(* IEC 61131-3 sources: ZPLC/conformance/cmp (part 2) *)

(* ---- cmp-020-two-enums-same-value-name.st ---- *)
TYPE A : (X, Y); END_TYPE
TYPE B : (Y, Z); END_TYPE

PROGRAM Main
VAR
  fromA AT %QW0 : INT;
  fromB AT %QW1 : INT;
  zB AT %QW2 : INT;
END_VAR
  fromA := A#Y;
  fromB := B#Y;
  zB := B#Z;
END_PROGRAM

(* ---- cmp-021-concat-leaves-its-arguments.st ---- *)
PROGRAM Main
VAR
  a : STRING[16] := 'ab';
  b : STRING[16] := 'cd';
  r : STRING[16];
  la AT %QW0 : INT;
  lb AT %QW1 : INT;
  lr AT %QW2 : INT;
  ok AT %QX6.0 : BOOL;
END_VAR
  r := CONCAT(a, b);
  la := LEN(a);
  lb := LEN(b);
  lr := LEN(r);
  ok := r = 'abcd';
END_PROGRAM

(* ---- cmp-021-find.st ---- *)
PROGRAM Main
VAR
  s : STRING[16] := 'HELLO';
  p1 AT %QW0 : INT;
  p2 AT %QW1 : INT;
  p3 AT %QW2 : INT;
  p4 AT %QW3 : INT;
END_VAR
  p1 := FIND(s, 'LL');
  p2 := FIND(s, 'H');
  p3 := FIND(s, 'LOL');
  p4 := FIND(s, 'O');
END_PROGRAM

(* ---- cmp-021-function-returning-a-string.st ---- *)
FUNCTION Tag : STRING[8]
VAR_INPUT n : INT; END_VAR
  IF n = 1 THEN
    Tag := 'one';
  ELSE
    Tag := 'other';
  END_IF;
END_FUNCTION

PROGRAM Main
VAR
  r : STRING[12];
  l AT %QW0 : INT;
  ok AT %QX2.0 : BOOL;
END_VAR
  r := CONCAT(Tag(1), Tag(2));
  l := LEN(r);
  ok := r = 'oneother';
END_PROGRAM

(* ---- cmp-021-initial-literal-longer-than-capacity-rejected.st ---- *)
PROGRAM Main
VAR
  s : STRING[3] := 'abcd';
END_VAR
END_PROGRAM

(* ---- cmp-021-insert-delete-replace.st ---- *)
PROGRAM Main
VAR
  s : STRING[16] := 'HELLO';
  i : STRING[16];
  d : STRING[16];
  r : STRING[16];
  ls AT %QW0 : INT;
  oki AT %QX2.0 : BOOL;
  okd AT %QX2.1 : BOOL;
  okr AT %QX2.2 : BOOL;
END_VAR
  i := INSERT(s, 'XY', 2);
  d := DELETE(s, 2, 2);
  r := REPLACE(s, 'AB', 2, 3);
  ls := LEN(s);
  oki := i = 'HEXYLLO';
  okd := d = 'HLO';
  okr := r = 'HABO';
END_PROGRAM

(* ---- cmp-021-left-and-right-beyond-the-length.st ---- *)
PROGRAM Main
VAR
  s : STRING[16] := 'abc';
  l : STRING[16];
  r : STRING[16];
  ll AT %QW0 : INT;
  lr AT %QW1 : INT;
  z AT %QW2 : INT;
END_VAR
  l := LEFT(s, 10);
  r := RIGHT(s, 10);
  ll := LEN(l);
  lr := LEN(r);
  z := LEN(LEFT(s, 0));
END_PROGRAM

(* ---- cmp-021-left-right-mid-keep-the-argument.st ---- *)
PROGRAM Main
VAR
  s : STRING[16] := 'HELLO';
  l : STRING[16];
  r : STRING[16];
  m : STRING[16];
  ls AT %QW0 : INT;
  okl AT %QX2.0 : BOOL;
  okr AT %QX2.1 : BOOL;
  okm AT %QX2.2 : BOOL;
END_VAR
  l := LEFT(s, 2);
  r := RIGHT(s, 3);
  m := MID(s, 2, 3);
  ls := LEN(s);
  okl := l = 'HE';
  okr := r = 'LLO';
  okm := m = 'ELL';
END_PROGRAM

(* ---- cmp-021-literal-longer-than-capacity-rejected.st ---- *)
PROGRAM Main
VAR
  s : STRING[3];
END_VAR
  s := 'abcd';
END_PROGRAM

(* ---- cmp-021-nested-string-functions.st ---- *)
PROGRAM Main
VAR
  a : STRING[16] := 'one';
  b : STRING[16] := 'two';
  r : STRING[16];
  l AT %QW0 : INT;
  ok AT %QX2.0 : BOOL;
  eq AT %QX2.1 : BOOL;
END_VAR
  r := CONCAT(LEFT(a, 2), RIGHT(b, 2));
  l := LEN(r);
  ok := r = 'onwo';
  eq := LEFT(a, 1) = LEFT('ozone', 1);
END_PROGRAM

(* ---- cmp-021-string-assign-length.st ---- *)
PROGRAM Text
VAR
  s : STRING;
  n AT %QW0 : INT;
END_VAR
  s := 'hello';
  n := LEN(s);
END_PROGRAM

(* ---- cmp-021-string-assignment-between-variables.st ---- *)
PROGRAM Main
VAR
  a : STRING[16];
  b : STRING[16];
  la AT %QW0 : INT;
  lb AT %QW1 : INT;
  same AT %QX4.0 : BOOL;
END_VAR
  a := 'hello';
  b := a;
  a := 'x';
  la := LEN(a);
  lb := LEN(b);
  same := b = 'hello';
END_PROGRAM

(* ---- cmp-021-string-buffer-survives-a-function-call.st ---- *)
FUNCTION Mark : INT
VAR_INPUT k : INT; END_VAR
  Mark := LEN(CONCAT('abc', 'defg')) + k;
END_FUNCTION

FUNCTION Pair : INT
VAR_INPUT
  x : STRING[8];
  m : INT;
END_VAR
  Pair := LEN(x) * 100 + m;
END_FUNCTION

PROGRAM Main
VAR
  a : STRING[8] := 'hello';
  r AT %QW0 : INT;
END_VAR
  r := Pair(LEFT(a, 2), Mark(1));
END_PROGRAM

(* ---- cmp-021-string-built-from-itself.st ---- *)
PROGRAM Main
VAR
  e : STRING[8] := 'AB';
  f : STRING[8] := 'AB';
  g : STRING[8] := 'ABCD';
  h : STRING[8] := 'ABCDE';
  okE AT %QX0.0 : BOOL;
  okF AT %QX0.1 : BOOL;
  okG AT %QX0.2 : BOOL;
  okH AT %QX0.3 : BOOL;
END_VAR
  e := CONCAT(e, e);
  f := CONCAT('xy', f);
  g := INSERT(g, '--', 2);
  h := REPLACE(h, 'Y', 2, 3);
  okE := e = 'ABAB';
  okF := f = 'xyAB';
  okG := g = 'AB--CD';
  okH := h = 'AYE';
END_PROGRAM

(* ---- cmp-021-string-comparison.st ---- *)
PROGRAM Main
VAR
  a : STRING[16] := 'abc';
  b : STRING[16] := 'abc';
  c : STRING[16] := 'abd';
  same AT %QX0.0 : BOOL;
  differ AT %QX0.1 : BOOL;
  literal AT %QX0.2 : BOOL;
END_VAR
  same := a = b;
  differ := a <> c;
  literal := c = 'abd';
END_PROGRAM

(* ---- cmp-021-string-cut-in-place.st ---- *)
PROGRAM Main
VAR
  a : STRING[8] := 'ABCDEFGH';
  b : STRING[8] := 'ABCDEFGH';
  c : STRING[8] := 'ABCDEFGH';
  d : STRING[8] := 'ABCDEFGH';
  okA AT %QX0.0 : BOOL;
  okB AT %QX0.1 : BOOL;
  okC AT %QX0.2 : BOOL;
  okD AT %QX0.3 : BOOL;
  lenA AT %QW1 : INT;
END_VAR
  a := LEFT(a, 3);
  b := RIGHT(b, 3);
  c := MID(c, 3, 2);
  d := DELETE(d, 3, 4);
  okA := a = 'ABC';
  okB := b = 'FGH';
  okC := c = 'CD';
  okD := d = 'ABGH';
  lenA := LEN(a);
END_PROGRAM

(* ---- cmp-021-string-function-into-array-element.st ---- *)
PROGRAM Main
VAR
  names : ARRAY[0..2] OF STRING[10];
  i : INT := 1;
  src : STRING[10] := 'pressure';
  l AT %QW0 : INT;
  ok AT %QX2.0 : BOOL;
END_VAR
  names[i] := LEFT(src, 4);
  l := LEN(names[1]);
  ok := names[1] = 'pres';
END_PROGRAM

(* ---- cmp-021-string-function-keeps-argument.st ---- *)
PROGRAM Text
VAR
  left AT %QW0 : INT;
  whole AT %QW1 : INT;
END_VAR
  left := LEN(LEFT('hello', 2));
  whole := LEN('hello');
END_PROGRAM

(* ---- cmp-021-string-function-reading-its-target-in-a-count.st ---- *)
PROGRAM Main
VAR
  k : STRING[8] := 'abcdef';
  t : STRING[8] := 'wxyz';
  okK AT %QX0.0 : BOOL;
  okT AT %QX0.1 : BOOL;
END_VAR
  k := LEFT(k, LEN(k) - 2);
  t := LEFT(t, LEN(k) - 1);
  okK := k = 'abcd';
  okT := t = 'wxy';
END_PROGRAM

(* ---- cmp-021-string-initial-values.st ---- *)
PROGRAM Main
VAR
  a : STRING := 'abc';
  b : STRING[10] := 'hi';
  c : STRING[16];
  la AT %QW0 : INT;
  lb AT %QW1 : INT;
  lc AT %QW2 : INT;
  ok AT %QX6.0 : BOOL;
END_VAR
  la := LEN(a);
  lb := LEN(b);
  lc := LEN(c);
  ok := b = 'hi';
END_PROGRAM

(* ---- cmp-021-string-literal-length.st ---- *)
PROGRAM Text
VAR
  n AT %QW0 : INT;
END_VAR
  n := LEN('hello');
END_PROGRAM

(* ---- cmp-021-string-members-and-elements.st ---- *)
TYPE Label : STRUCT id : INT; text : STRING[12]; END_STRUCT END_TYPE

PROGRAM Main
VAR
  l : Label;
  a : ARRAY[0..1] OF STRING[8];
  lt AT %QW0 : INT;
  la AT %QW1 : INT;
  id AT %QW2 : INT;
  ok AT %QX6.0 : BOOL;
END_VAR
  l.id := 42;
  l.text := 'motor 1';
  a[1] := 'pump';
  lt := LEN(l.text);
  la := LEN(a[1]);
  id := l.id;
  ok := a[1] = 'pump';
END_PROGRAM

(* ---- cmp-021-string-parameter-is-a-copy.st ---- *)
FUNCTION Shout : INT
VAR_INPUT text : STRING[16]; END_VAR
  text := CONCAT(text, '!');
  Shout := LEN(text);
END_FUNCTION

PROGRAM Main
VAR
  s : STRING[16] := 'hello';
  inside AT %QW0 : INT;
  outside AT %QW1 : INT;
END_VAR
  inside := Shout(s);
  outside := LEN(s);
END_PROGRAM

(* ---- cmp-021-string-truncates-to-its-capacity.st ---- *)
PROGRAM Main
VAR
  long : STRING[16] := 'abcdefgh';
  short : STRING[5];
  l AT %QW0 : INT;
  ok AT %QX2.0 : BOOL;
END_VAR
  short := long;
  l := LEN(short);
  ok := short = 'abcde';
END_PROGRAM

(* ---- cmp-021-string-with-capacity.st ---- *)
PROGRAM Text
VAR
  s : STRING[20];
  n AT %QW0 : INT;
END_VAR
  s := 'hello';
  n := LEN(s);
END_PROGRAM

(* ---- cmp-021-wstring-assignment.st ---- *)
PROGRAM Main
VAR
  a : WSTRING[10] := "hi";
  b : WSTRING[10];
  la AT %QW0 : INT;
  lb AT %QW1 : INT;
END_VAR
  b := "world";
  la := LEN(a);
  lb := LEN(b);
  a := b;
  la := LEN(a) * 10 + la;
END_PROGRAM

(* ---- cmp-021-wstring-literal-length.st ---- *)
PROGRAM WideLiteral
VAR
  n AT %QW0 : INT;
END_VAR
  n := LEN("abcd");
END_PROGRAM

(* ---- cmp-021-wstring-variable-length.st ---- *)
PROGRAM WideVariable
VAR
  w : WSTRING := "abcd";
  n AT %QW0 : INT;
END_VAR
  n := LEN(w);
END_PROGRAM

(* ---- cmp-022-array-bound-constant-expression.st ---- *)
VAR_GLOBAL CONSTANT N : INT := 2; END_VAR

PROGRAM Main
VAR
  a : ARRAY[N - 2 .. N * 2 - 1] OF INT;
  last AT %QW0 : INT;
END_VAR
  a[3] := 33;
  last := a[3];
END_PROGRAM

(* ---- cmp-022-array-constant-bound.st ---- *)
VAR_GLOBAL CONSTANT N : INT := 4; END_VAR

PROGRAM Table
VAR
  a : ARRAY[0..N] OF INT;
  last AT %QW0 : INT;
END_VAR
  a[4] := 9;
  last := a[4];
END_PROGRAM

(* ---- cmp-022-array-element-read-write.st ---- *)
PROGRAM Table
VAR
  a : ARRAY[1..4] OF INT;
  i : INT;
  third AT %QW0 : INT;
END_VAR
  FOR i := 1 TO 4 DO
    a[i] := i * 10;
  END_FOR;
  third := a[3];
END_PROGRAM

(* ---- cmp-022-array-index-from-array.st ---- *)
PROGRAM Main
VAR
  b : ARRAY[0..2] OF INT;
  a : ARRAY[0..4] OF DINT;
  v AT %QD0 : DINT;
END_VAR
  b[1] := 4;
  a[4] := 654321;
  v := a[b[1]];
END_PROGRAM

(* ---- cmp-022-array-initialiser-large-repeat.st ---- *)
PROGRAM Main
VAR
  a : ARRAY[0..99] OF INT := [100(3)];
  first AT %QW0 : INT;
  last AT %QW1 : INT;
  after AT %QW2 : INT;
END_VAR
  first := a[0];
  last := a[99];
  after := a[50] + 4;
END_PROGRAM

(* ---- cmp-022-array-initialiser-list.st ---- *)
PROGRAM Table
VAR
  a : ARRAY[0..2] OF INT := [1, 2, 3];
  seen AT %QW0 : INT;
END_VAR
  seen := a[1];
END_PROGRAM

(* ---- cmp-022-array-initialiser-of-structures.st ---- *)
TYPE Pt : STRUCT x : INT; z : DINT; END_STRUCT END_TYPE

PROGRAM Main
VAR
  a : ARRAY[0..1] OF Pt := [(x := 1, z := 100000), (x := 2, z := 200000)];
  x1 AT %QW0 : INT;
  z0 AT %QD1 : DINT;
  z1 AT %QD2 : DINT;
END_VAR
  x1 := a[1].x;
  z0 := a[0].z;
  z1 := a[1].z;
END_PROGRAM

(* ---- cmp-022-array-initialiser-repeat.st ---- *)
PROGRAM Table
VAR
  a : ARRAY[0..3] OF INT := [4(7)];
  seen AT %QW0 : INT;
END_VAR
  seen := a[3];
END_PROGRAM

(* ---- cmp-022-array-initialiser-two-dimensions.st ---- *)
PROGRAM Main
VAR
  a : ARRAY[0..1, 0..2] OF INT := [[1, 2, 3], [4, 5, 6]];
  b : ARRAY[0..1, 0..1] OF INT := [10, 20, 30, 40];
  mid AT %QW0 : INT;
  last AT %QW1 : INT;
  flat AT %QW2 : INT;
END_VAR
  mid := a[1, 1];
  last := a[1, 2];
  flat := b[1, 0];
END_PROGRAM

(* ---- cmp-022-array-inside-structure.st ---- *)
TYPE Rec : STRUCT n : INT; a : ARRAY[1..3] OF DINT; tail : INT; END_STRUCT END_TYPE

PROGRAM Main
VAR
  s : Rec;
  i : INT;
  second AT %QD0 : DINT;
  tail AT %QW2 : INT;
END_VAR
  s.tail := 77;
  FOR i := 1 TO 3 DO
    s.a[i] := i * 100000;
  END_FOR;
  second := s.a[2];
  tail := s.tail;
END_PROGRAM

(* ---- cmp-022-array-negative-lower-bound.st ---- *)
PROGRAM Table
VAR
  a : ARRAY[-5..5] OF INT;
  total AT %QW0 : INT;
END_VAR
  a[-5] := 3;
  a[0] := 4;
  total := a[-5] + a[0];
END_PROGRAM

(* ---- cmp-022-array-of-lint-negative.st ---- *)
PROGRAM Main
VAR
  a : ARRAY[0..3] OF LINT;
  b : LINT;
  same AT %QX0.0 : BOOL;
  negative AT %QX0.1 : BOOL;
  neighbour AT %QX0.2 : BOOL;
END_VAR
  a[1] := -5;
  a[2] := 7;
  b := a[1];
  same := a[1] = -5;
  negative := b < 0;
  neighbour := a[2] = 7;
END_PROGRAM

(* ---- cmp-022-array-of-lint-variable-index.st ---- *)
PROGRAM Main
VAR
  a : ARRAY[0..3] OF LINT;
  i : INT := 2;
  big : LINT := 5000000000;
  back : LINT;
  same AT %QX0.0 : BOOL;
  other AT %QX0.1 : BOOL;
  low AT %QD1 : DINT;
END_VAR
  a[i] := big;
  a[i + 1] := -9;
  back := a[i];
  same := back = 5000000000;
  other := a[3] = -9;
  low := a[2] - 5000000000;
END_PROGRAM

(* ---- cmp-022-array-of-lint.st ---- *)
PROGRAM Table
VAR
  a : ARRAY[0..3] OF LINT;
  ok AT %QX0.0 : BOOL;
END_VAR
  a[2] := 1;
  ok := a[2] = 1;
END_PROGRAM

(* ---- cmp-022-array-of-real-and-bool.st ---- *)
PROGRAM Main
VAR
  r : ARRAY[0..2] OF REAL;
  f : ARRAY[0..2] OF BOOL;
  sum AT %QD0 : REAL;
  second AT %QX4.0 : BOOL;
  third AT %QX4.1 : BOOL;
END_VAR
  r[0] := 1.5;
  r[1] := 2.25;
  r[2] := 0.25;
  f[1] := TRUE;
  sum := r[0] + r[1] + r[2];
  second := f[1];
  third := f[2];
END_PROGRAM

(* ---- cmp-022-array-of-structures-index-expression.st ---- *)
TYPE Pt : STRUCT x : INT; z : DINT; END_STRUCT END_TYPE

PROGRAM Main
VAR
  a : ARRAY[0..3] OF Pt;
  i : INT;
  z2 AT %QD0 : DINT;
  x3 AT %QW2 : INT;
  x0 AT %QW3 : INT;
END_VAR
  FOR i := 0 TO 3 DO
    a[i].z := i * 1000 + 70000;
    a[i].x := -i;
  END_FOR;
  z2 := a[2].z;
  x3 := a[3].x;
  x0 := a[0].x;
END_PROGRAM

(* ---- cmp-022-array-of-structures.st ---- *)
TYPE Pt : STRUCT x : INT; y : INT; z : DINT; END_STRUCT END_TYPE

PROGRAM Table
VAR
  a : ARRAY[0..3] OF Pt;
  seen AT %QW0 : INT;
END_VAR
  a[1].x := 5;
  seen := a[1].x;
END_PROGRAM

(* ---- cmp-022-array-two-dimensions-negative-bounds.st ---- *)
PROGRAM Main
VAR
  a : ARRAY[-1..1, 0..2] OF INT;
  r : INT;
  c : INT;
  low AT %QW0 : INT;
  high AT %QW1 : INT;
  mid AT %QW2 : INT;
END_VAR
  FOR r := -1 TO 1 DO
    FOR c := 0 TO 2 DO
      a[r, c] := r * 10 + c;
    END_FOR;
  END_FOR;
  low := a[-1, 2];
  high := a[1, 0];
  mid := a[0, 1];
END_PROGRAM

(* ---- cmp-022-multi-dimensional-arrays.st ---- *)
PROGRAM Grid
VAR
  plane : ARRAY[0..1, 0..2] OF INT;
  cube : ARRAY[1..2, 1..2, 1..2] OF DINT;
  gains : ARRAY[0..2] OF REAL;
  flags : ARRAY[0..3] OF BOOL;
  i : INT;
  j : INT;
  corner AT %QW0 : INT;
  inner AT %QW1 : INT;
  far AT %QD1 : DINT;
  gain AT %QD2 : REAL;
  flag AT %QX12.0 : BOOL;
  clear AT %QX12.1 : BOOL;
END_VAR
  FOR i := 0 TO 1 DO
    FOR j := 0 TO 2 DO
      plane[i, j] := i * 10 + j;
    END_FOR;
  END_FOR;
  cube[2, 1, 2] := 212;
  gains[2] := 1.5;
  flags[3] := TRUE;
  corner := plane[1, 2];
  inner := plane[0, 1];
  far := cube[2, 1, 2];
  gain := gains[2];
  flag := flags[3];
  clear := flags[0];
END_PROGRAM

(* ---- cmp-023-array-index-out-of-bounds-faults.st ---- *)
PROGRAM Table
VAR
  a : ARRAY[0..1] OF INT;
  index : INT := 2;
END_VAR
  a[index] := 77;
END_PROGRAM

(* ---- cmp-023-constant-index-in-second-dimension-rejected.st ---- *)
PROGRAM Main
VAR
  a : ARRAY[0..1, 0..2] OF INT;
  v AT %QW0 : INT;
END_VAR
  v := a[1, 3];
END_PROGRAM

(* ---- cmp-023-constant-index-out-of-bounds.st ---- *)
PROGRAM Table
VAR
  a : ARRAY[0..3] OF INT;
END_VAR
  a[10] := 1;
END_PROGRAM

(* ---- cmp-023-index-at-both-bounds-is-accepted.st ---- *)
PROGRAM Main
VAR
  a : ARRAY[2..4] OF INT;
  i : INT;
  first AT %QW0 : INT;
  last AT %QW1 : INT;
END_VAR
  i := 2;
  a[i] := 12;
  i := 4;
  a[i] := 14;
  i := 2;
  first := a[i];
  i := 4;
  last := a[i];
END_PROGRAM

(* ---- cmp-023-index-below-lower-bound-faults.st ---- *)
PROGRAM Main
VAR
  a : ARRAY[2..4] OF INT;
  i : INT := 1;
END_VAR
  a[i] := 5;
END_PROGRAM

(* ---- cmp-023-negative-constant-index-rejected.st ---- *)
PROGRAM Main
VAR
  a : ARRAY[0..3] OF INT;
END_VAR
  a[-1] := 1;
END_PROGRAM

(* ---- cmp-023-read-out-of-bounds-faults.st ---- *)
PROGRAM Main
VAR
  a : ARRAY[0..3] OF DINT;
  i : INT := 4;
  v AT %QD0 : DINT;
END_VAR
  v := a[i];
END_PROGRAM

(* ---- cmp-023-second-dimension-out-of-bounds-faults.st ---- *)
PROGRAM Main
VAR
  a : ARRAY[0..1, 0..2] OF INT;
  j : INT := 3;
  v AT %QW0 : INT;
END_VAR
  v := a[1, j];
END_PROGRAM

(* ---- cmp-024-dereference-of-non-reference-rejected.st ---- *)
PROGRAM Main
VAR
  x : INT;
  y : INT;
END_VAR
  y := x^;
END_PROGRAM

(* ---- cmp-024-null-reference-faults.st ---- *)
PROGRAM Pointer
VAR
  p : REF_TO INT;
  seen AT %QW0 : INT;
END_VAR
  seen := p^;
END_PROGRAM

(* ---- cmp-024-ref-of-another-type.st ---- *)
PROGRAM Pointer
VAR
  r : REAL;
  p : REF_TO INT;
END_VAR
  p := REF(r);
END_PROGRAM

(* ---- cmp-024-ref-to-reads-and-writes-the-referenced-variable.st ---- *)
PROGRAM Reference
VAR
  target : INT := 5;
  link : REF_TO INT;
  seen AT %QW0 : INT;
  moved AT %QW1 : INT;
END_VAR
  link := REF(target);
  seen := link^;
  link^ := 42;
  moved := target;
END_PROGRAM

(* ---- cmp-024-reference-is-null-until-assigned.st ---- *)
PROGRAM Main
VAR
  x : INT;
  p : REF_TO INT;
  before AT %QX0.0 : BOOL;
  after AT %QX0.1 : BOOL;
END_VAR
  before := p = NULL;
  p := REF(x);
  after := p = NULL;
END_PROGRAM

(* ---- cmp-024-reference-of-wrong-type-passed-rejected.st ---- *)
FUNCTION Peek : INT
VAR_INPUT r : REF_TO INT; END_VAR
  Peek := r^;
END_FUNCTION

PROGRAM Main
VAR
  d : DINT;
  seen AT %QW0 : INT;
END_VAR
  seen := Peek(REF(d));
END_PROGRAM

(* ---- cmp-024-reference-of-wrong-type-variable-rejected.st ---- *)
PROGRAM Main
VAR
  d : DINT;
  p : REF_TO INT;
END_VAR
  p := REF(d);
END_PROGRAM

(* ---- cmp-024-reference-passed-to-a-function.st ---- *)
FUNCTION Peek : INT
VAR_INPUT r : REF_TO INT; END_VAR
  Peek := r^;
END_FUNCTION

PROGRAM Main
VAR
  v : INT := 41;
  seen AT %QW0 : INT;
END_VAR
  seen := Peek(REF(v)) + 1;
END_PROGRAM

(* ---- cmp-024-reference-read-and-write.st ---- *)
PROGRAM Main
VAR
  x : INT;
  p : REF_TO INT;
  seen AT %QW0 : INT;
  direct AT %QW1 : INT;
END_VAR
  p := REF(x);
  p^ := 7;
  seen := p^;
  direct := x;
END_PROGRAM

(* ---- cmp-024-reference-stored-in-a-number-rejected.st ---- *)
PROGRAM Main
VAR
  d : DINT;
  e : DINT;
END_VAR
  d := REF(e);
END_PROGRAM

(* ---- cmp-024-reference-to-a-structure.st ---- *)
TYPE Pt : STRUCT x : INT; z : DINT; END_STRUCT END_TYPE

PROGRAM Main
VAR
  s : Pt;
  pp : REF_TO Pt;
  x AT %QW0 : INT;
  z AT %QD1 : DINT;
END_VAR
  pp := REF(s);
  pp^.z := 123456;
  pp^.x := -7;
  x := s.x;
  z := pp^.z;
END_PROGRAM

(* ---- cmp-024-reference-to-member-and-element.st ---- *)
TYPE Pt : STRUCT x : INT; z : DINT; END_STRUCT END_TYPE

PROGRAM Main
VAR
  s : Pt;
  a : ARRAY[0..3] OF DINT;
  pz : REF_TO DINT;
  pe : REF_TO DINT;
  z AT %QD0 : DINT;
  e2 AT %QD1 : DINT;
END_VAR
  pz := REF(s.z);
  pz^ := 123456;
  pe := REF(a[2]);
  pe^ := 654321;
  z := s.z;
  e2 := a[2];
END_PROGRAM

(* ---- cmp-025-fifo-default-size-is-eight.st ---- *)
PROGRAM DefaultQueue
VAR
  push AT %IX0.0 : BOOL;
  item AT %ID1 : DINT;
  line : FIFO;
  count AT %QD0 : DINT;
  full AT %QX4.0 : BOOL;
END_VAR
  line(PUSH := push, DATA_IN := item);
  count := line.COUNT;
  full := line.FULL;
END_PROGRAM

(* ---- cmp-025-function-local-initial-value.st ---- *)
FUNCTION Offset : INT
VAR_INPUT a : INT; END_VAR
VAR k : INT := 100; END_VAR
  Offset := a + k;
END_FUNCTION

PROGRAM Locals
VAR
  seen AT %QW0 : INT;
END_VAR
  seen := Offset(1);
END_PROGRAM

(* ---- cmp-025-global-initial-value.st ---- *)
VAR_GLOBAL G : INT := 42; END_VAR

PROGRAM Globals
VAR
  seen AT %QW0 : INT;
END_VAR
  seen := G;
END_PROGRAM

(* ---- cmp-025-global-structure-and-array-initial-values.st ---- *)
TYPE Pt : STRUCT x : INT := 3; z : DINT := 90000; END_STRUCT END_TYPE

VAR_GLOBAL
  g : Pt;
  t : ARRAY[0..2] OF INT := [4, 5, 6];
END_VAR

PROGRAM Main
VAR
  x AT %QW0 : INT;
  z AT %QD1 : DINT;
  t2 AT %QW4 : INT;
END_VAR
  x := g.x;
  z := g.z;
  t2 := t[2];
END_PROGRAM

(* ---- cmp-025-initial-value-is-written-once.st ---- *)
PROGRAM Main
VAR
  n : INT := 5;
  seen AT %QW0 : INT;
END_VAR
  n := n + 1;
  seen := n;
END_PROGRAM

(* ---- cmp-025-initial-values-of-each-type.st ---- *)
PROGRAM Main
VAR
  flag : BOOL := TRUE;
  ratio : REAL := 1.5;
  big : DINT := -70000;
  wait : TIME := T#2s;
  oflag AT %QX0.0 : BOOL;
  oratio AT %QD1 : REAL;
  obig AT %QD2 : DINT;
  owait AT %QD3 : TIME;
END_VAR
  oflag := flag;
  oratio := ratio;
  obig := big;
  owait := wait;
END_PROGRAM

(* ---- cmp-025-lifo-default-size-is-eight.st ---- *)
PROGRAM DefaultStack
VAR
  push AT %IX0.0 : BOOL;
  item AT %ID1 : DINT;
  pile : LIFO;
  count AT %QD0 : DINT;
  full AT %QX4.0 : BOOL;
END_VAR
  pile(PUSH := push, DATA_IN := item);
  count := pile.COUNT;
  full := pile.FULL;
END_PROGRAM

(* ---- cmp-026-assignment-to-a-constant.st ---- *)
VAR_GLOBAL CONSTANT K : INT := 42; END_VAR

PROGRAM Constants
VAR
  x : INT;
END_VAR
  K := 3;
  x := K;
END_PROGRAM

(* ---- cmp-026-constants-of-real-and-integer.st ---- *)
VAR_GLOBAL CONSTANT
  HALF : REAL := 0.5;
  STEP : INT := 4;
END_VAR

PROGRAM Main
VAR
  r AT %QD0 : REAL;
  n AT %QW2 : INT;
END_VAR
  r := HALF * 3.0;
  n := STEP * 3;
END_PROGRAM

(* ---- cmp-026-global-constant-value.st ---- *)
VAR_GLOBAL CONSTANT K : INT := 42; END_VAR

PROGRAM Constants
VAR
  seen AT %QW0 : INT;
END_VAR
  seen := K;
END_PROGRAM

(* ---- cmp-026-var-constant-assignment-rejected.st ---- *)
PROGRAM Main
VAR CONSTANT
  K : INT := 5;
END_VAR
VAR
  x : INT;
END_VAR
  K := 6;
  x := K;
END_PROGRAM

(* ---- cmp-026-var-constant.st ---- *)
PROGRAM Constants
VAR CONSTANT
  K : INT := 5;
END_VAR
VAR
  seen AT %QW0 : INT;
END_VAR
  seen := K;
END_PROGRAM

(* ---- cmp-027-function-local-initial-value-on-every-call.st ---- *)
FUNCTION Step : INT
VAR_INPUT x : INT; END_VAR
VAR k : INT := 10; END_VAR
  k := k + x;
  Step := k;
END_FUNCTION

PROGRAM Main
VAR
  first AT %QW0 : INT;
  second AT %QW1 : INT;
END_VAR
  first := Step(1);
  second := Step(2);
END_PROGRAM

(* ---- cmp-027-function-local-not-retained.st ---- *)
FUNCTION Count : INT
VAR_INPUT x : INT; END_VAR
VAR k : INT; END_VAR
  k := k + 1;
  Count := k;
END_FUNCTION

PROGRAM Calls
VAR
  first AT %QW0 : INT;
  second AT %QW1 : INT;
END_VAR
  first := Count(0);
  second := Count(0);
END_PROGRAM

(* ---- cmp-027-function-local-string-and-array.st ---- *)
FUNCTION Grow : INT
VAR_INPUT n : INT; END_VAR
VAR
  s : STRING[16];
  a : ARRAY[0..2] OF INT;
END_VAR
  a[1] := a[1] + n;
  s := CONCAT(s, 'ab');
  Grow := LEN(s) * 10 + a[1];
END_FUNCTION

PROGRAM Main
VAR
  r AT %QW0 : INT;
END_VAR
  r := Grow(3);
END_PROGRAM

(* ---- cmp-029-non-retain-accepted.st ---- *)
PROGRAM Volatile
VAR NON_RETAIN
  count : INT;
END_VAR
VAR
  seen AT %QW0 : INT;
END_VAR
  count := count + 1;
  seen := count;
END_PROGRAM

(* ---- cmp-029-retain-and-ordinary-variables-together.st ---- *)
PROGRAM Mixed
VAR RETAIN
  kept : DINT;
  flag : BOOL;
END_VAR
VAR
  plain : INT;
  seen AT %QD0 : DINT;
  mark AT %QX4.0 : BOOL;
END_VAR
  kept := kept + 10;
  flag := kept > 15;
  plain := plain + 1;
  seen := kept + plain;
  mark := flag;
END_PROGRAM

(* ---- cmp-029-retain-global-with-initial-value.st ---- *)
VAR_GLOBAL RETAIN
  total : INT := 10;
END_VAR

PROGRAM Totals
VAR
  seen AT %QW0 : INT;
END_VAR
  total := total + 1;
  seen := total;
END_PROGRAM

(* ---- cmp-029-retain-structure-and-string.st ---- *)
TYPE Pair : STRUCT a : INT := 3; b : INT := 4; END_STRUCT END_TYPE

PROGRAM Mixed
VAR RETAIN
  p : Pair;
  s : STRING[10] := 'abc';
  n : INT := 2;
END_VAR
VAR
  sum AT %QW0 : INT;
  len AT %QW2 : INT;
END_VAR
  n := n + 1;
  sum := p.a + p.b + n;
  len := LEN(s);
END_PROGRAM

(* ---- cmp-029-var-global-retain.st ---- *)
VAR_GLOBAL RETAIN
  total : INT;
END_VAR

PROGRAM Totals
VAR
  seen AT %QW0 : INT;
END_VAR
  total := total + 2;
  seen := total;
END_PROGRAM

(* ---- cmp-029-var-non-retain-is-accepted.st ---- *)
PROGRAM Volatile
VAR NON_RETAIN
  x : INT := 5;
END_VAR
VAR
  q AT %QW0 : INT;
END_VAR
  q := x;
END_PROGRAM

(* ---- cmp-029-var-retain-accepted.st ---- *)
PROGRAM Retained
VAR RETAIN
  count : INT;
END_VAR
VAR
  seen AT %QW0 : INT;
END_VAR
  count := count + 1;
  seen := count;
END_PROGRAM

(* ---- cmp-030-alias-default-value.st ---- *)
TYPE Limit : INT := 100; END_TYPE

PROGRAM Defaults
VAR
  a : Limit;
  b : Limit := 7;
  sum AT %QW0 : INT;
END_VAR
  sum := a + b;
END_PROGRAM

(* ---- cmp-030-alias-of-array-and-structure.st ---- *)
TYPE
  Point : STRUCT x : INT; y : INT; END_STRUCT;
  Marker : Point;
  Samples : ARRAY[0..2] OF INT;
END_TYPE

PROGRAM Aliases
VAR
  m : Marker;
  s : Samples;
  total AT %QW0 : INT;
END_VAR
  m.x := 2;
  m.y := 3;
  s[0] := 10;
  s[2] := 20;
  total := m.x + m.y + s[0] + s[2];
END_PROGRAM

(* ---- cmp-030-alias-refers-to-itself.st ---- *)
TYPE A : B; B : A; END_TYPE

PROGRAM Cycle
VAR
  x : A;
END_VAR
END_PROGRAM

(* ---- cmp-030-function-var-output.st ---- *)
FUNCTION Twice : INT
VAR_INPUT a : INT; END_VAR
VAR_OUTPUT o : INT; END_VAR
  o := a;
  Twice := a + a;
END_FUNCTION

PROGRAM Outputs
VAR
  seen AT %QW0 : INT;
END_VAR
  seen := Twice(3);
END_PROGRAM

(* ---- cmp-030-several-names-one-declaration.st ---- *)
PROGRAM Names
VAR
  a, b : INT;
  total AT %QW0 : INT;
END_VAR
  a := 3;
  b := 4;
  total := a + b;
END_PROGRAM

(* ---- cmp-030-several-names-with-initial-value.st ---- *)
PROGRAM Names
VAR
  a, b, c : INT := 4;
  total AT %QW0 : INT;
END_VAR
  total := a + b + c;
END_PROGRAM

(* ---- cmp-030-several-types-one-block.st ---- *)
TYPE
  A : STRUCT v : INT; END_STRUCT;
  B : (R, G);
END_TYPE

PROGRAM Types
VAR
  a : A;
  seen AT %QW0 : INT;
END_VAR
  a.v := 6;
  seen := a.v;
END_PROGRAM

(* ---- cmp-030-type-alias.st ---- *)
TYPE MyInt : INT; END_TYPE

PROGRAM Alias
VAR
  x : MyInt;
  seen AT %QW0 : INT;
END_VAR
  x := 9;
  seen := x;
END_PROGRAM

(* ---- cmp-030-var-external-type-differs.st ---- *)
VAR_GLOBAL G : INT; END_VAR

PROGRAM External
VAR_EXTERNAL G : REAL; END_VAR
VAR
  seen AT %QW0 : INT;
END_VAR
  seen := 1;
END_PROGRAM

(* ---- cmp-030-var-external-without-global.st ---- *)
PROGRAM External
VAR_EXTERNAL Missing : INT; END_VAR
VAR
  seen AT %QW0 : INT;
END_VAR
  seen := Missing;
END_PROGRAM

(* ---- cmp-030-var-external.st ---- *)
VAR_GLOBAL G : INT; END_VAR

PROGRAM External
VAR_EXTERNAL G : INT; END_VAR
VAR
  seen AT %QW0 : INT;
END_VAR
  G := 5;
  seen := G;
END_PROGRAM

(* ---- cmp-030-var-temp-in-program.st ---- *)
PROGRAM Temporary
VAR_TEMP
  k : INT;
END_VAR
VAR
  seen AT %QW0 : INT;
END_VAR
  k := 6;
  seen := k;
END_PROGRAM

(* ---- cmp-031-0x-form-still-works.st ---- *)
PROGRAM Literal
VAR
  seen AT %QW0 : INT;
END_VAR
  seen := 0xFF;
END_PROGRAM

(* ---- cmp-031-base-not-supported.st ---- *)
PROGRAM Literal
VAR
  seen AT %QW0 : INT;
END_VAR
  seen := 3#12;
END_PROGRAM

(* ---- cmp-031-binary-literal.st ---- *)
PROGRAM Literal
VAR
  seen AT %QW0 : INT;
END_VAR
  seen := 2#1010;
END_PROGRAM

(* ---- cmp-031-c-style-hexadecimal-keeps-working.st ---- *)
PROGRAM CStyle
VAR
  n AT %QW0 : INT;
END_VAR
  n := 0xFF;
END_PROGRAM

(* ---- cmp-031-digit-separator.st ---- *)
PROGRAM Literal
VAR
  seen AT %QW0 : INT;
END_VAR
  seen := 1_000;
END_PROGRAM

(* ---- cmp-031-hexadecimal-literal.st ---- *)
PROGRAM Literal
VAR
  seen AT %QW0 : INT;
END_VAR
  seen := 16#FF;
END_PROGRAM

(* ---- cmp-031-negative-based-literal.st ---- *)
PROGRAM Literal
VAR
  seen AT %QW0 : INT;
END_VAR
  seen := -16#10;
END_PROGRAM

(* ---- cmp-031-octal-literal.st ---- *)
PROGRAM Octal
VAR
  n AT %QW0 : INT;
END_VAR
  n := 8#17;
END_PROGRAM

(* ---- cmp-031-separator-in-based-literal.st ---- *)
PROGRAM Literal
VAR
  seen AT %QW0 : INT;
END_VAR
  seen := 2#1111_0000;
END_PROGRAM

(* ---- cmp-031-typed-literal-out-of-range.st ---- *)
PROGRAM Literal
VAR
  seen AT %QW0 : INT;
END_VAR
  seen := SINT#200;
END_PROGRAM

(* ---- cmp-031-typed-literal.st ---- *)
PROGRAM Literal
VAR
  seen AT %QW0 : INT;
END_VAR
  seen := INT#5;
END_PROGRAM

(* ---- cmp-031-typed-literals-of-each-kind.st ---- *)
PROGRAM Literal
VAR
  small AT %QW0 : INT;
  bits AT %QD2 : DWORD;
  flag AT %QX6.0 : BOOL;
  half AT %QD8 : REAL;
END_VAR
  small := SINT#-3 + INT#4;
  bits := DWORD#16#DEAD_BEEF;
  flag := BOOL#TRUE;
  half := REAL#1.5;
END_PROGRAM

(* ---- cmp-032-ampersand-binds-tighter-than-or.st ---- *)
PROGRAM Logic
VAR
  a : BOOL := TRUE;
  b : BOOL := FALSE;
  c : BOOL := FALSE;
  seen AT %QX0.0 : BOOL;
END_VAR
  seen := a OR b & c;
END_PROGRAM

(* ---- cmp-032-ampersand-operator.st ---- *)
PROGRAM Both
VAR
  a : BOOL := TRUE;
  b : BOOL := TRUE;
  both AT %QX0.0 : BOOL;
END_VAR
  both := a & b;
END_PROGRAM

(* ---- cmp-032-bit-access-of-bool-rejected.st ---- *)
PROGRAM Bits
VAR
  f : BOOL;
  seen AT %QX0.0 : BOOL;
END_VAR
  seen := f.0;
END_PROGRAM

(* ---- cmp-032-bit-access.st ---- *)
PROGRAM Bits
VAR
  w : WORD := 1;
  low AT %QX0.0 : BOOL;
END_VAR
  low := w.0;
END_PROGRAM

(* ---- cmp-032-bit-number-out-of-range.st ---- *)
PROGRAM Bits
VAR
  b : BYTE;
  seen AT %QX0.0 : BOOL;
END_VAR
  seen := b.8;
END_PROGRAM

(* ---- cmp-032-bit-of-lword.st ---- *)
PROGRAM Bits
VAR
  l : LWORD;
  low AT %QX0.0 : BOOL;
  high AT %QX0.1 : BOOL;
  other AT %QX0.2 : BOOL;
END_VAR
  l.40 := TRUE;
  low := l.0;
  high := l.40;
  other := l.39;
END_PROGRAM

(* ---- cmp-032-bit-of-member-and-element.st ---- *)
TYPE Status : STRUCT flags : WORD; END_STRUCT END_TYPE

PROGRAM Bits
VAR
  s : Status;
  a : ARRAY[0..1] OF WORD;
  one AT %QX0.0 : BOOL;
  two AT %QX0.1 : BOOL;
END_VAR
  s.flags := 16#0004;
  a[1] := 16#0100;
  one := s.flags.2;
  a[1].0 := TRUE;
  two := a[1].8 AND a[1].0;
END_PROGRAM

(* ---- cmp-032-bit-set-and-clear.st ---- *)
PROGRAM Bits
VAR
  w AT %QW0 : WORD;
END_VAR
  w := 0;
  w.3 := TRUE;
  w.0 := TRUE;
  w.3 := FALSE;
  w.15 := TRUE;
END_PROGRAM

(* ---- cmp-032-bit-write-in-each-width.st ---- *)
PROGRAM Bits
VAR
  b AT %QB0 : BYTE;
  i AT %QW2 : INT;
  d AT %QD4 : DWORD;
END_VAR
  b.7 := TRUE;
  i.15 := TRUE;
  d.31 := TRUE;
  d.0 := TRUE;
END_PROGRAM

(* ---- cmp-032-block-comment.st ---- *)
PROGRAM Comment
VAR
  seen AT %QW0 : INT;
END_VAR
  /* a comment */ seen := 1;
END_PROGRAM

(* ---- cmp-032-comment-delimiters-inside-comments.st ---- *)
PROGRAM Comments
VAR
  seen AT %QW0 : INT;
END_VAR
  (* a /* inside *) seen := 1;
  /* a (* inside */ seen := seen + 1;
  // (* not an opener
  seen := seen + 1; /* trailing */ (* and another *)
END_PROGRAM

(* ---- cmp-032-empty-statement.st ---- *)
PROGRAM Empty
VAR
  seen AT %QW0 : INT;
END_VAR
  seen := 1;;
END_PROGRAM

(* ---- cmp-032-empty-statements-inside-blocks.st ---- *)
PROGRAM Empty
VAR
  seen AT %QW0 : INT;
END_VAR
  ;
  IF TRUE THEN ; seen := 2;; END_IF;;
  CASE seen OF 2: ; seen := seen + 1; END_CASE;
END_PROGRAM

(* ---- cmp-032-exponent-operator.st ---- *)
PROGRAM Power
VAR
  cube AT %QD0 : REAL;
END_VAR
  cube := 2.0 ** 3.0;
END_PROGRAM

(* ---- cmp-032-power-fractional-exponent.st ---- *)
PROGRAM Power
VAR
  d1 : REAL;
  d2 : REAL;
  d3 : REAL;
  d4 : REAL;
  root AT %QX0.0 : BOOL;
  cube AT %QX0.1 : BOOL;
  big AT %QX0.2 : BOOL;
  small AT %QX0.3 : BOOL;
END_VAR
  d1 := 9.0 ** 0.5 - 3.0;
  d2 := 27.0 ** (1.0 / 3.0) - 3.0;
  d3 := 10.0 ** 2.5 / 316.227766 - 1.0;
  d4 := 0.5 ** 1.5 / 0.35355339 - 1.0;
  root := (d1 < 0.0001) AND (d1 > -0.0001);
  cube := (d2 < 0.0001) AND (d2 > -0.0001);
  big := (d3 < 0.00005) AND (d3 > -0.00005);
  small := (d4 < 0.00005) AND (d4 > -0.00005);
END_PROGRAM

(* ---- cmp-032-power-negative-and-zero-exponent.st ---- *)
PROGRAM Power
VAR
  r AT %QD0 : REAL;
  s AT %QD4 : REAL;
  t AT %QD8 : REAL;
END_VAR
  r := 2.0 ** -2.0;
  s := 5.0 ** 0.0;
  t := 0.0 ** 0.0;
END_PROGRAM

(* ---- cmp-032-power-negative-base.st ---- *)
PROGRAM Power
VAR
  r AT %QD0 : REAL;
  s AT %QD4 : REAL;
END_VAR
  r := (-3.0) ** 3.0;
  s := (-2.0) ** 2.0;
END_PROGRAM

(* ---- cmp-032-power-of-integers.st ---- *)
PROGRAM Power
VAR
  a : INT := 2;
  r AT %QD0 : REAL;
  s AT %QD4 : REAL;
END_VAR
  r := 2 ** 10;
  s := a ** 3;
END_PROGRAM

(* ---- cmp-032-power-precedence.st ---- *)
PROGRAM Power
VAR
  r AT %QD0 : REAL;
  s AT %QD4 : REAL;
END_VAR
  r := -2.0 ** 2.0;
  s := 2.0 * 3.0 ** 2.0;
END_PROGRAM

(* ---- cmp-032-power-zero-base-negative-exponent-faults.st ---- *)
PROGRAM Power
VAR
  zero : REAL := 0.0;
  r AT %QD0 : REAL;
END_VAR
  r := zero ** -1.0;
END_PROGRAM

(* ---- cmp-033-library-block-in-lower-case.st ---- *)
PROGRAM Timer
VAR
  t : ton;
  done AT %QX0.0 : BOOL;
END_VAR
  t(IN := TRUE, PT := T#20ms);
  done := t.Q;
END_PROGRAM

(* ---- cmp-033-library-block-name-as-variable.st ---- *)
PROGRAM Names
VAR
  Pulse : BOOL;
  seen AT %QX0.0 : BOOL;
END_VAR
  Pulse := TRUE;
  seen := Pulse;
END_PROGRAM

(* ---- cmp-034-function-does-not-see-a-program-variable.st ---- *)
FUNCTION Peek : INT
VAR_INPUT n : INT; END_VAR
  Peek := n + hidden;
END_FUNCTION

PROGRAM Scopes
VAR
  hidden : INT := 5;
  out AT %QW0 : INT;
END_VAR
  out := Peek(1);
END_PROGRAM

(* ---- cmp-034-function-locals-do-not-clash.st ---- *)
FUNCTION Pick : INT
VAR_INPUT a : INT; b : INT; END_VAR
VAR tmp : INT; END_VAR
  tmp := a;
  Pick := tmp + b;
END_FUNCTION

FUNCTION Mix : INT
VAR_INPUT b : INT; a : INT; END_VAR
VAR tmp : INT; END_VAR
  tmp := a * 10;
  Mix := tmp + b;
END_FUNCTION

PROGRAM Scopes
VAR
  a : INT := 1000;
  tmp : INT := 2000;
  first AT %QW0 : INT;
  second AT %QW1 : INT;
  kept AT %QW2 : INT;
END_VAR
  first := Pick(1, 2);
  second := Mix(1, 2);
  kept := a + tmp;
END_PROGRAM

(* ---- cmp-034-function-reads-a-global.st ---- *)
VAR_GLOBAL
  base : INT := 100;
END_VAR

FUNCTION Offset : INT
VAR_INPUT n : INT; END_VAR
VAR_EXTERNAL base : INT; END_VAR
  Offset := n + base;
END_FUNCTION

PROGRAM Scopes
VAR
  out AT %QW0 : INT;
  other AT %QW1 : INT;
END_VAR
  out := Offset(5);
  other := Offset(n := 6);
END_PROGRAM

(* ---- cmp-034-function-with-loops-and-locals-of-the-same-name.st ---- *)
FUNCTION SumTo : DINT
VAR_INPUT n : INT; END_VAR
VAR i : INT; total : DINT; END_VAR
  FOR i := 1 TO n DO
    total := total + i;
  END_FOR;
  SumTo := total;
END_FUNCTION

FUNCTION SumSquares : DINT
VAR_INPUT n : INT; END_VAR
VAR i : INT; total : DINT; END_VAR
  FOR i := 1 TO n DO
    total := total + i * i;
  END_FOR;
  SumSquares := total;
END_FUNCTION

PROGRAM Loops
VAR
  i : INT := 100;
  total : DINT := 1000;
  sum AT %QD0 : DINT;
  squares AT %QD1 : DINT;
  again AT %QD2 : DINT;
  program_i AT %QW6 : INT;
END_VAR
  sum := SumTo(4);
  squares := SumSquares(3);
  again := SumTo(4);
  program_i := i;
END_PROGRAM

(* ---- cmp-034-parameter-shadows-program-variable.st ---- *)
FUNCTION Succ : INT
VAR_INPUT a : INT; END_VAR
  Succ := a + 1;
END_FUNCTION

PROGRAM Scopes
VAR
  a : INT := 9;
  total AT %QW0 : INT;
END_VAR
  total := Succ(1) + a;
END_PROGRAM

(* ---- cmp-034-same-parameter-name-two-functions.st ---- *)
FUNCTION Succ : INT
VAR_INPUT a : INT; END_VAR
  Succ := a + 1;
END_FUNCTION

FUNCTION Twice : INT
VAR_INPUT a : INT; END_VAR
  Twice := a * 2;
END_FUNCTION

PROGRAM Scopes
VAR
  total AT %QW0 : INT;
END_VAR
  total := Succ(1) + Twice(2);
END_PROGRAM

(* ---- cmp-035-call-statement-runs-the-function.st ---- *)
VAR_GLOBAL
  counter : INT;
END_VAR

FUNCTION Bump : INT
VAR_INPUT amount : INT; END_VAR
VAR_EXTERNAL counter : INT; END_VAR
  counter := counter + amount;
  Bump := counter;
END_FUNCTION

PROGRAM Statement
VAR
  seen AT %QW0 : INT;
END_VAR
  Bump(2);
  Bump(amount := 3);
  seen := counter;
END_PROGRAM

(* ---- cmp-035-function-call-as-statement.st ---- *)
FUNCTION Succ : INT
VAR_INPUT a : INT; END_VAR
  Succ := a + 1;
END_FUNCTION

PROGRAM Statement
VAR
  seen AT %QW0 : INT;
END_VAR
  Succ(1);
  seen := 5;
END_PROGRAM

(* ---- cmp-035-missing-argument.st ---- *)
FUNCTION Sub : INT
VAR_INPUT a : INT; b : INT; END_VAR
  Sub := a - b;
END_FUNCTION

PROGRAM Arguments
VAR
  x : INT;
END_VAR
  x := Sub(10);
END_PROGRAM

(* ---- cmp-035-named-arguments-any-order.st ---- *)
FUNCTION Sub : INT
VAR_INPUT a : INT; b : INT; END_VAR
  Sub := a - b;
END_FUNCTION

PROGRAM Arguments
VAR
  diff AT %QW0 : INT;
END_VAR
  diff := Sub(b := 1, a := 10);
END_PROGRAM

(* ---- cmp-035-parameter-given-twice-is-rejected.st ---- *)
FUNCTION Sub : INT
VAR_INPUT a : INT; b : INT; END_VAR
  Sub := a - b;
END_FUNCTION

PROGRAM Arguments
VAR
  x : INT;
END_VAR
  x := Sub(1, a := 2, b := 3);
END_PROGRAM

(* ---- cmp-035-parameter-with-a-declared-value-may-be-left-out.st ---- *)
FUNCTION Scale : INT
VAR_INPUT value : INT; factor : INT := 10; END_VAR
  Scale := value * factor;
END_FUNCTION

PROGRAM Arguments
VAR
  by_default AT %QW0 : INT;
  given AT %QW1 : INT;
END_VAR
  by_default := Scale(3);
  given := Scale(3, 2);
END_PROGRAM

(* ---- cmp-035-positional-after-named-is-rejected.st ---- *)
FUNCTION Sub : INT
VAR_INPUT a : INT; b : INT; END_VAR
  Sub := a - b;
END_FUNCTION

PROGRAM Arguments
VAR
  x : INT;
END_VAR
  x := Sub(a := 1, 2);
END_PROGRAM

(* ---- cmp-035-positional-then-named.st ---- *)
FUNCTION Sub3 : INT
VAR_INPUT a : INT; b : INT; c : INT; END_VAR
  Sub3 := a - b - c;
END_FUNCTION

PROGRAM Arguments
VAR
  mixed AT %QW0 : INT;
  named AT %QW1 : INT;
END_VAR
  mixed := Sub3(10, c := 1, b := 2);
  named := Sub3(c := 1, a := 10, b := 2);
END_PROGRAM

(* ---- cmp-035-recursion-through-two-functions.st ---- *)
FUNCTION Ping : INT
VAR_INPUT n : INT; END_VAR
  IF n > 0 THEN
    Ping := Pong(n - 1);
  END_IF;
END_FUNCTION

FUNCTION Pong : INT
VAR_INPUT n : INT; END_VAR
  Pong := Ping(n);
END_FUNCTION

PROGRAM Recursion
VAR
  x : INT;
END_VAR
  x := Ping(3);
END_PROGRAM

(* ---- cmp-035-recursive-call.st ---- *)
FUNCTION Fact : INT
VAR_INPUT n : INT; END_VAR
  IF n <= 1 THEN
    Fact := 1;
  ELSE
    Fact := n * Fact(n - 1);
  END_IF;
END_FUNCTION

PROGRAM Recursion
VAR
  x : INT;
END_VAR
  x := Fact(5);
END_PROGRAM

(* ---- cmp-035-too-many-arguments-is-rejected.st ---- *)
FUNCTION Sub : INT
VAR_INPUT a : INT; b : INT; END_VAR
  Sub := a - b;
END_FUNCTION

PROGRAM Arguments
VAR
  x : INT;
END_VAR
  x := Sub(1, 2, 3);
END_PROGRAM

(* ---- cmp-035-unknown-argument-name.st ---- *)
FUNCTION Sub : INT
VAR_INPUT a : INT; b : INT; END_VAR
  Sub := a - b;
END_FUNCTION

PROGRAM Arguments
VAR
  x : INT;
END_VAR
  x := Sub(a := 1, c := 2);
END_PROGRAM

(* ---- cmp-036-return-in-a-program-ends-its-scan.st ---- *)
PROGRAM Returns
VAR
  x AT %QW0 : INT;
END_VAR
  x := 1;
  RETURN;
  x := 2;
END_PROGRAM

(* ---- cmp-036-return-leaves-the-function-only.st ---- *)
FUNCTION Clamp : INT
VAR_INPUT a : INT; END_VAR
  Clamp := a;
  IF a > 10 THEN
    Clamp := 10;
    RETURN;
  END_IF;
END_FUNCTION

PROGRAM Returns
VAR
  clamped AT %QW0 : INT;
  after AT %QX2.0 : BOOL;
END_VAR
  clamped := Clamp(50);
  after := TRUE;
END_PROGRAM

(* ---- cmp-037-input-bound-with-arrow-is-rejected.st ---- *)
PROGRAM Binding
VAR
  t : TON;
  seen : BOOL;
END_VAR
  t(IN => seen, PT := T#10ms);
END_PROGRAM

(* ---- cmp-037-output-binding.st ---- *)
PROGRAM Binding
VAR
  t : TON;
  done AT %QX0.0 : BOOL;
END_VAR
  t(IN := TRUE, PT := T#10ms, Q => done);
END_PROGRAM

(* ---- cmp-037-unknown-parameter-standard-block.st ---- *)
PROGRAM Timer
VAR
  t : TON;
END_VAR
  t(IN := TRUE, PT := T#10ms, BOGUS := 5);
END_PROGRAM

(* ---- cmp-038-array-of-instances.st ---- *)
PROGRAM Composition
VAR
  timers : ARRAY[0..1] OF TON;
  done AT %QX0.0 : BOOL;
END_VAR
  timers[0](IN := TRUE, PT := T#10ms);
  done := timers[0].Q;
END_PROGRAM

(* ---- cmp-038-array-run-time-index.st ---- *)
PROGRAM Counters
VAR
  c : ARRAY[0..2] OF CTU;
  i : INT;
  first AT %QW0 : INT;
  second AT %QW2 : INT;
  third AT %QW4 : INT;
END_VAR
  c[i](CU := TRUE, PV := 100);
  i := i + 1;
  IF i > 2 THEN i := 0; END_IF;
  first := c[0].CV;
  second := c[1].CV;
  third := c[2].CV;
END_PROGRAM

(* ---- cmp-038-constant-index-out-of-bounds.st ---- *)
PROGRAM Composition
VAR
  t : ARRAY[0..1] OF TON;
END_VAR
  t[2](IN := TRUE, PT := T#10ms);
END_PROGRAM

(* ---- cmp-039-continue-skips-the-rest-of-the-body.st ---- *)
PROGRAM Skipping
VAR
  i : INT;
  total AT %QW0 : INT;
  passes AT %QW1 : INT;
END_VAR
  FOR i := 1 TO 6 DO
    passes := passes + 1;
    IF i MOD 2 = 0 THEN
      CONTINUE;
    END_IF;
    total := total + i;
  END_FOR;
END_PROGRAM

(* ---- cmp-039-for-counting-down.st ---- *)
PROGRAM Loop
VAR
  i : INT;
  steps AT %QW0 : INT;
END_VAR
  steps := 0;
  FOR i := 3 TO 1 BY -1 DO
    steps := steps + 1;
  END_FOR;
END_PROGRAM

(* ---- cmp-039-for-variable-negative-step.st ---- *)
PROGRAM Loop
VAR
  i : DINT;
  step : DINT := -2;
  steps AT %QW0 : INT;
END_VAR
  steps := 0;
  FOR i := 6 TO 1 BY step DO
    steps := steps + 1;
  END_FOR;
END_PROGRAM

(* ---- cmp-039-repeat-until.st ---- *)
PROGRAM Loop
VAR
  i : INT;
  seen AT %QW0 : INT;
END_VAR
  i := 0;
  REPEAT
    i := i + 1;
  UNTIL i >= 3
  END_REPEAT;
  seen := i;
END_PROGRAM

(* ---- cmp-039-while-and-exit.st ---- *)
PROGRAM Loop
VAR
  i : INT;
  seen AT %QW0 : INT;
END_VAR
  i := 0;
  WHILE TRUE DO
    i := i + 1;
    IF i >= 5 THEN
      EXIT;
    END_IF;
  END_WHILE;
  seen := i;
END_PROGRAM

(* ---- cmp-040-case-enum-label.st ---- *)
TYPE St : (IDLE, RUN); END_TYPE

PROGRAM Select
VAR
  state : St;
  picked AT %QW0 : INT;
END_VAR
  state := RUN;
  CASE state OF
    IDLE: picked := 1;
    RUN: picked := 2;
  END_CASE;
END_PROGRAM

(* ---- cmp-040-case-integer-list.st ---- *)
PROGRAM Select
VAR
  i : INT := 2;
  picked AT %QW0 : INT;
END_VAR
  CASE i OF
    1: picked := 10;
    2, 3: picked := 20;
  ELSE
    picked := 30;
  END_CASE;
END_PROGRAM

(* ---- cmp-040-case-negative-label.st ---- *)
PROGRAM Select
VAR
  i : DINT := -1;
  picked AT %QW0 : INT;
END_VAR
  CASE i OF
    -1: picked := 1;
  ELSE
    picked := 2;
  END_CASE;
END_PROGRAM

(* ---- cmp-040-case-range.st ---- *)
PROGRAM Select
VAR
  i : INT := 3;
  picked AT %QW0 : INT;
END_VAR
  CASE i OF
    1..5: picked := 1;
  ELSE
    picked := 2;
  END_CASE;
END_PROGRAM

(* ---- cmp-040-case-without-else-in-a-loop.st ---- *)
PROGRAM CaseLoop
VAR
  i : INT;
  hits : INT;
  total AT %QW0 : INT;
END_VAR
  hits := 0;
  FOR i := 1 TO 10 DO
    CASE i OF
      3: hits := hits + 1;
      7: hits := hits + 10;
    END_CASE;
  END_FOR;
  total := hits;
END_PROGRAM

(* ---- cmp-040-overlapping-case-labels.st ---- *)
PROGRAM Select
VAR
  i : INT;
  picked : INT;
END_VAR
  CASE i OF
    1, 2: picked := 1;
    2, 3: picked := 2;
  END_CASE;
END_PROGRAM

(* ---- cmp-042-debug-map-addresses-of-every-program-consumer.st ---- *)
PROGRAM Consumer
VAR
  consumed : INT;
  small : BYTE;
END_VAR
  consumed := Shared + 1;
  small := 7;
END_PROGRAM

(* ---- cmp-042-debug-map-addresses-of-every-program.st ---- *)
PROGRAM Producer
VAR
  produced : INT;
  total : DINT;
  ratio : REAL;
  tag : STRING[12];
  gate : Gate;
END_VAR
  produced := 11;
  total := 100000;
  ratio := 2.5;
  tag := 'unit';
  gate(open := TRUE);
  Shared := 44;
END_PROGRAM

(* ---- cmp-042-function-block-declared-in-two-files-is-rejected.st ---- *)
PROGRAM Project
END_PROGRAM

(* ---- cmp-042-function-block-in-another-file.st ---- *)
PROGRAM Project
VAR
  d : Echo;
  seen AT %QX0.0 : BOOL;
END_VAR
  d(sig := TRUE);
  seen := d.out;
END_PROGRAM

(* ---- cmp-042-function-from-another-file-in-two-programs-right.st ---- *)
PROGRAM Right
VAR
  r AT %QW1 : INT;
END_VAR
  r := Twice(x := 5) + 1;
END_PROGRAM

(* ---- cmp-042-function-from-another-file-in-two-programs.st ---- *)
PROGRAM Left
VAR
  r AT %QW0 : INT;
END_VAR
  r := Twice(x := 4);
END_PROGRAM

(* ---- cmp-042-global-in-another-file.st ---- *)
PROGRAM Project
VAR
  seen AT %QW0 : INT;
END_VAR
  Shared := 7;
  seen := Shared;
END_PROGRAM

(* ---- cmp-042-global-initial-value-is-applied-once-bump.st ---- *)
PROGRAM Bumper
VAR
  scans AT %QW1 : INT;
END_VAR
  Counter := Counter + 1;
  scans := scans + 1;
END_PROGRAM

(* ---- cmp-042-global-initial-value-is-applied-once.st ---- *)
PROGRAM Reader
VAR
  seen AT %QW0 : INT;
END_VAR
  seen := Counter;
END_PROGRAM

(* ---- cmp-042-two-tasks-share-a-global-reader.st ---- *)
PROGRAM Reader
VAR
  seen AT %QW1 : INT;
END_VAR
  seen := Shared;
END_PROGRAM

(* ---- cmp-042-two-tasks-share-a-global.st ---- *)
PROGRAM Writer
VAR
  mine AT %QW0 : INT;
END_VAR
  Shared := 7;
  mine := Shared;
END_PROGRAM

(* ---- cmp-042-type-from-another-file-in-a-structure.st ---- *)
TYPE Segment : STRUCT
  a : Point;
  b : Point;
END_STRUCT END_TYPE

PROGRAM Geometry
VAR
  s : Segment;
  total AT %QW0 : INT;
END_VAR
  s.a.x := 3;
  s.a.y := 4;
  s.b.x := 10;
  s.b.y := 20;
  total := s.a.x + s.a.y + s.b.x + s.b.y;
END_PROGRAM

(* ---- cmp-043-allocation-failure-states-bytes-and-consumers.st ---- *)
PROGRAM Overflow
VAR
  Table : ARRAY[0..8999] OF BYTE;
  Gain : REAL;
END_VAR
  Gain := 1.5;
END_PROGRAM

(* ---- cmp-043-array-beyond-256-bytes.st ---- *)
PROGRAM Large
VAR
  a : ARRAY[0..199] OF INT;
  last AT %QW0 : INT;
END_VAR
  a[199] := 7;
  last := a[199];
END_PROGRAM

(* ---- cmp-043-program-that-fills-the-region.st ---- *)
PROGRAM Fill
VAR
  all : ARRAY[0..8190] OF BYTE;
  seen AT %QW0 : INT;
END_VAR
  all[0] := 1;
  all[8190] := 2;
  seen := all[0] + all[8190];
END_PROGRAM

(* ---- cmp-043-programs-share-the-region-second.st ---- *)
PROGRAM Second
VAR
  block : ARRAY[0..299] OF BYTE;
  seen AT %QW1 : INT;
END_VAR
  block[299] := 9;
  seen := block[299];
END_PROGRAM

(* ---- cmp-043-programs-share-the-region.st ---- *)
PROGRAM First
VAR
  block : ARRAY[0..299] OF BYTE;
  seen AT %QW0 : INT;
END_VAR
  block[299] := 5;
  seen := block[299];
END_PROGRAM

(* ---- cmp-043-three-strings.st ---- *)
PROGRAM Large
VAR
  a : STRING;
  b : STRING;
  c : STRING;
  seen AT %QW0 : INT;
END_VAR
  seen := 1;
END_PROGRAM

(* ---- cmp-044-located-memory-overlap.st ---- *)
PROGRAM Overlap
VAR
  a AT %MW0 : INT;
  b : INT;
END_VAR
  b := a;
END_PROGRAM

(* ---- cmp-044-located-memory-variable.st ---- *)
PROGRAM Marker
VAR
  m AT %MW0 : INT;
  out AT %QW0 : INT;
END_VAR
  m := m + 1;
  out := m;
END_PROGRAM

(* ---- cmp-047-direct-addresses-of-every-width.st ---- *)
PROGRAM Widths
VAR
  in_bit AT %IX0.3 : BOOL;
  in_byte AT %IB1 : BYTE;
  in_word AT %IW1 : WORD;
  in_dword AT %ID1 : DWORD;
  out_bit AT %QX0.5 : BOOL;
  out_byte AT %QB1 : BYTE;
  out_word AT %QW1 : WORD;
  out_dword AT %QD1 : DWORD;
END_VAR
  out_bit := in_bit;
  out_byte := in_byte;
  out_word := in_word;
  out_dword := in_dword;
END_PROGRAM

(* ---- cmp-047-two-cyclic-tasks-of-one-interval-right.st ---- *)
PROGRAM Right
VAR
  runs AT %QW1 : INT;
END_VAR
  runs := runs + 1;
END_PROGRAM

(* ---- cmp-047-two-cyclic-tasks-of-one-interval.st ---- *)
PROGRAM Left
VAR
  runs AT %QW0 : INT;
END_VAR
  runs := runs + 1;
END_PROGRAM

(* ---- cmp-047-two-programs-writing-one-output-are-rejected-second.st ---- *)
PROGRAM Second
VAR
  motor AT %QX0.0 : BOOL;
END_VAR
  motor := FALSE;
END_PROGRAM

(* ---- cmp-047-two-programs-writing-one-output-are-rejected.st ---- *)
PROGRAM First
VAR
  motor AT %QX0.0 : BOOL;
END_VAR
  motor := TRUE;
END_PROGRAM

(* ---- cmp-049-direct-address-beyond-the-operand-field-is-rejected.st ---- *)
PROGRAM Main
VAR
  far AT %MW40000 : INT;
END_VAR
far := 1;
END_PROGRAM

(* ---- cmp-050-expression-too-deep-for-the-stack-is-rejected.st ---- *)
PROGRAM Main
VAR
  a : DINT := 1;
  r AT %QD0 : DINT;
END_VAR
r := a + (a + (a + (a + (a + (a + (a + (a + (a + (a + (a + (a + (a + (a + (a + (a + (a + (a + (a + (a + (a + (a + (a + (a + (a + (a + (a + (a + (a + (a + (a + (a + (a + (a + (a + (a + (a + (a + (a + (a + (a + (a + (a + (a + (a + (a + (a + (a + (a + (a + (a + (a + (a + (a + (a + (a + (a + (a + (a + (a + (a + (a + (a + (a + (a + (a + (a + (a + (a + (a + (a + (a + (a + (a + (a + (a + (a + (a + (a + (a + (a + (a + (a + (a + (a + (a + (a + (a + (a + (a + (a + (a + (a + (a + (a + (a + (a + (a + (a + (a + (a + (a + (a + (a + (a + (a + (a + (a + (a + (a + (a + (a + (a + (a + (a + (a + (a + (a + (a + (a + (a + (a + (a + (a + (a + (a + (a + (a + (a + (a + (a + (a + (a + (a + (a + (a + (a + (a + (a + (a)))))))))))))))))))))))))))))))))))))))))))))))))))))))))))))))))))))))))))))))))))))))))))))))))))))))))))))))))))))))))))))))))))))))))));
END_PROGRAM

(* ---- cmp-054-debug-map-address-with-a-type.st ---- *)
TYPE Pt : STRUCT x : INT; y : INT; END_STRUCT END_TYPE

PROGRAM Mapped
VAR
  p : Pt;
  s : INT;
  copy AT %QW0 : INT;
END_VAR
  s := 42;
  copy := s;
END_PROGRAM

(* ---- cmp-054-debug-map-lists-a-global.st ---- *)
VAR_GLOBAL G : INT; END_VAR

PROGRAM Mapped
VAR
  seen AT %QW0 : INT;
END_VAR
  G := 9;
  seen := G;
END_PROGRAM

(* ---- cmp-057-bool-and-round-conversions.st ---- *)
PROGRAM Conversions
VAR
  truth : BOOL := TRUE;
  zero : INT := 0;
  five : INT := 5;
  low : REAL := 2.4;
  high : REAL := 2.6;
  below : REAL := -2.6;
  as_int AT %QW0 : INT;
  from_zero AT %QX2.0 : BOOL;
  from_five AT %QX2.1 : BOOL;
  rounded_low AT %QD2 : REAL;
  rounded_high AT %QD3 : REAL;
  rounded_below AT %QD4 : REAL;
END_VAR
  as_int := BOOL_TO_INT(truth);
  from_zero := INT_TO_BOOL(zero);
  from_five := INT_TO_BOOL(five);
  rounded_low := ROUND(low);
  rounded_high := ROUND(high);
  rounded_below := ROUND(below);
END_PROGRAM

(* ---- cmp-057-conversions-to-bool-and-from-bool.st ---- *)
PROGRAM Booleans
VAR
  zero : REAL := 0.0;
  half : REAL := 0.5;
  minus_two : REAL := -2.0;
  minus_one : REAL := -1.0;
  big : REAL := 1.0E38;
  neg_zero : REAL;
  inf : REAL;
  nan : REAL;
  minus_int : INT := -1;
  high_only : DWORD := 16#10000;
  none : USINT := 0;
  yes : BOOL := TRUE;
  q0 AT %QX0.0 : BOOL;
  q1 AT %QX0.1 : BOOL;
  q2 AT %QX0.2 : BOOL;
  q3 AT %QX0.3 : BOOL;
  q4 AT %QX0.4 : BOOL;
  q5 AT %QX0.5 : BOOL;
  q6 AT %QX0.6 : BOOL;
  q7 AT %QX0.7 : BOOL;
  b0 AT %QB1 : USINT;
  b1 AT %QW1 : INT;
  b2 AT %QD1 : DINT;
END_VAR
  neg_zero := zero * minus_one;
  inf := big * big;
  nan := inf - inf;
  q0 := REAL_TO_BOOL(zero);
  q1 := REAL_TO_BOOL(half);
  q2 := REAL_TO_BOOL(minus_two);
  q3 := REAL_TO_BOOL(neg_zero);
  q4 := INT_TO_BOOL(minus_int);
  q5 := DWORD_TO_BOOL(high_only);
  q6 := USINT_TO_BOOL(none);
  q7 := REAL_TO_BOOL(nan);
  b0 := BOOL_TO_USINT(yes);
  b1 := BOOL_TO_INT(yes);
  b2 := BOOL_TO_DINT(yes);
END_PROGRAM

(* ---- cmp-057-dint-to-real-exists.st ---- *)
PROGRAM Convert
VAR
  n : DINT := 100000;
  r AT %QD0 : REAL;
END_VAR
  r := DINT_TO_REAL(n);
END_PROGRAM

(* ---- cmp-057-int-to-dint-exists.st ---- *)
PROGRAM Convert
VAR
  n : INT := 7;
  d AT %QD0 : DINT;
END_VAR
  d := INT_TO_DINT(n);
END_PROGRAM

(* ---- cmp-057-integer-conversion-functions.st ---- *)
PROGRAM Conversions
VAR
  small : SINT := -3;
  half : INT := -300;
  whole : DINT := -70000;
  unsigned_half : UINT := 65535;
  octet : BYTE := 200;
  word_value : WORD := 40000;
  a AT %QW0 : INT;
  b AT %QW1 : INT;
  c AT %QD1 : DINT;
  d AT %QD2 : DINT;
  e AT %QW8 : INT;
  f AT %QD3 : DINT;
END_VAR
  a := SINT_TO_INT(small);
  b := DINT_TO_INT(half);
  c := INT_TO_DINT(half);
  d := UINT_TO_DINT(unsigned_half);
  e := BYTE_TO_INT(octet);
  f := WORD_TO_DINT(word_value);
END_PROGRAM

(* ---- cmp-057-integer-conversions-wrap-to-the-destination-width.st ---- *)
PROGRAM Wrap
VAR
  big : INT := 300;
  wide : DINT := 70000;
  max_uint : UINT := 65535;
  minus_one : INT := -1;
  minus_sint : SINT := -1;
  all_ones : UDINT := 4294967295;
  dword_value : DWORD := 16#12345678;
  word_value : WORD := 16#ABCD;
  r0 AT %QB0 : SINT;
  r1 AT %QW1 : INT;
  r2 AT %QW2 : INT;
  r3 AT %QB6 : USINT;
  r4 AT %QW4 : UINT;
  r5 AT %QW5 : UINT;
  r6 AT %QD3 : UDINT;
  r7 AT %QD4 : DINT;
  r8 AT %QW10 : WORD;
  r9 AT %QB22 : BYTE;
  r10 AT %QB23 : BYTE;
  r11 AT %QW12 : INT;
END_VAR
  r0 := INT_TO_SINT(big);
  r1 := DINT_TO_INT(wide);
  r2 := UINT_TO_INT(max_uint);
  r3 := INT_TO_USINT(minus_one);
  r4 := INT_TO_UINT(minus_one);
  r5 := SINT_TO_UINT(minus_sint);
  r6 := INT_TO_UDINT(minus_one);
  r7 := UDINT_TO_DINT(all_ones);
  r8 := DWORD_TO_WORD(dword_value);
  r9 := DWORD_TO_BYTE(dword_value);
  r10 := WORD_TO_BYTE(word_value);
  r11 := WORD_TO_INT(word_value);
END_PROGRAM

(* ---- cmp-057-integer-types-convert-to-real.st ---- *)
PROGRAM ToReal
VAR
  s : SINT := -3;
  us : USINT := 200;
  ui : UINT := 60000;
  d : DINT := -70000;
  ud : UDINT := 3000000000;
  w : WORD := 40000;
  dw : DWORD := 16#80000000;
  b : BYTE := 255;
  t : BOOL := TRUE;
  r0 AT %QD0 : REAL;
  r1 AT %QD1 : REAL;
  r2 AT %QD2 : REAL;
  r3 AT %QD3 : REAL;
  r4 AT %QD4 : REAL;
  r5 AT %QD5 : REAL;
  r6 AT %QD6 : REAL;
  r7 AT %QD7 : REAL;
  r8 AT %QD8 : REAL;
END_VAR
  r0 := SINT_TO_REAL(s);
  r1 := USINT_TO_REAL(us);
  r2 := UINT_TO_REAL(ui);
  r3 := DINT_TO_REAL(d);
  r4 := UDINT_TO_REAL(ud);
  r5 := WORD_TO_REAL(w);
  r6 := DWORD_TO_REAL(dw);
  r7 := BYTE_TO_REAL(b);
  r8 := BOOL_TO_REAL(t);
END_PROGRAM

(* ---- cmp-057-real-to-int-rounds.st ---- *)
PROGRAM Convert
VAR
  r : REAL := 3.7;
  i AT %QW0 : INT;
END_VAR
  i := REAL_TO_INT(r);
END_PROGRAM

(* ---- cmp-057-real-to-int-ties-go-to-even.st ---- *)
PROGRAM Ties
VAR
  half : REAL := 0.5;
  one_half : REAL := 1.5;
  two_half : REAL := 2.5;
  three_half : REAL := 3.5;
  minus_half : REAL := -0.5;
  minus_one_half : REAL := -1.5;
  minus_two_half : REAL := -2.5;
  almost_half : REAL := 0.49999997;
  last_tie : REAL := 8388607.5;
  r0 AT %QW0 : INT;
  r1 AT %QW1 : INT;
  r2 AT %QW2 : INT;
  r3 AT %QW3 : INT;
  r4 AT %QW4 : INT;
  r5 AT %QW5 : INT;
  r6 AT %QW6 : INT;
  r7 AT %QW7 : INT;
  r8 AT %QD4 : DINT;
END_VAR
  r0 := REAL_TO_INT(half);
  r1 := REAL_TO_INT(one_half);
  r2 := REAL_TO_INT(two_half);
  r3 := REAL_TO_INT(three_half);
  r4 := REAL_TO_INT(minus_half);
  r5 := REAL_TO_INT(minus_one_half);
  r6 := REAL_TO_INT(minus_two_half);
  r7 := REAL_TO_INT(almost_half);
  r8 := REAL_TO_DINT(last_tie);
END_PROGRAM

(* ---- cmp-057-real-to-integer-saturates-at-the-destination-range.st ---- *)
PROGRAM Saturate
VAR
  inf_source : REAL := 1.0E38;
  inf : REAL;
  nan : REAL;
  q0 AT %QB0 : SINT;
  q1 AT %QB1 : SINT;
  q2 AT %QB2 : USINT;
  q3 AT %QB3 : USINT;
  q4 AT %QW2 : INT;
  q5 AT %QW3 : INT;
  q6 AT %QW4 : UINT;
  q7 AT %QD3 : UDINT;
  q8 AT %QD4 : UDINT;
  q9 AT %QD5 : DINT;
  q10 AT %QD6 : DINT;
  q11 AT %QD7 : UDINT;
END_VAR
  inf := inf_source * inf_source;
  nan := inf - inf;
  q0 := REAL_TO_SINT(200.0);
  q1 := REAL_TO_SINT(-200.0);
  q2 := REAL_TO_USINT(300.0);
  q3 := REAL_TO_USINT(-5.0);
  q4 := REAL_TO_INT(40000.0);
  q5 := REAL_TO_INT(-40000.0);
  q6 := REAL_TO_UINT(70000.0);
  q7 := REAL_TO_UDINT(5.0E9);
  q8 := REAL_TO_UDINT(3.0E9);
  q9 := REAL_TO_DINT(nan);
  q10 := REAL_TO_DINT(0.0 - inf);
  q11 := REAL_TO_UDINT(inf);
END_PROGRAM

(* ---- cmp-057-round-half-away-from-zero-and-large-values.st ---- *)
PROGRAM Round
VAR
  below_half : REAL := 0.49999997;
  two_half : REAL := 2.5;
  large : REAL := 3.0E9;
  r0 AT %QD0 : REAL;
  r1 AT %QD1 : REAL;
  r2 AT %QD2 : REAL;
  r3 AT %QD3 : REAL;
  r4 AT %QD4 : REAL;
END_VAR
  r0 := ROUND(below_half);
  r1 := ROUND(two_half);
  r2 := ROUND(0.0 - two_half);
  r3 := ROUND(large);
  r4 := ROUND(0.5);
END_PROGRAM

(* ---- cmp-057-time-conversions.st ---- *)
PROGRAM TimeValues
VAR
  after : TIME := T#1s500ms;
  q0 AT %QD0 : DINT;
  q1 AT %QD1 : TIME;
  q2 AT %QD2 : UDINT;
  q3 AT %QD3 : REAL;
  q4 AT %QD4 : TIME;
  q5 AT %QW10 : WORD;
END_VAR
  q0 := TIME_TO_DINT(T#2s);
  q1 := DINT_TO_TIME(1500);
  q2 := TIME_TO_UDINT(T#1h);
  q3 := TIME_TO_REAL(after);
  q4 := REAL_TO_TIME(2500.0);
  q5 := TIME_TO_WORD(T#70s);
END_PROGRAM

(* ---- cmp-057-tof-elapsed-stops-at-preset.st ---- *)
PROGRAM Delay
VAR
  n : INT;
  t : TOF;
  q AT %QX0.0 : BOOL;
  elapsed AT %QD1 : TIME;
END_VAR
  n := n + 1;
  t(IN := n <= 2, PT := T#50ms);
  q := t.Q;
  elapsed := t.ET;
END_PROGRAM

(* ---- cmp-057-ton-elapsed-stops-at-preset.st ---- *)
PROGRAM Timer
VAR
  t : TON;
  elapsed AT %QD0 : TIME;
END_VAR
  t(IN := TRUE, PT := T#50ms);
  elapsed := t.ET;
END_PROGRAM

(* ---- cmp-057-ton-zero-preset-follows-the-input.st ---- *)
PROGRAM Delay
VAR
  enable AT %IX0.0 : BOOL;
  t : TON;
  q AT %QX0.0 : BOOL;
END_VAR
  t(IN := enable, PT := T#0ms);
  q := t.Q;
END_PROGRAM

(* ---- cmp-057-tp-elapsed-resets-when-the-pulse-ends-with-input-low.st ---- *)
PROGRAM Pulse
VAR
  trigger AT %IX0.0 : BOOL;
  shot : TP;
  q AT %QX0.0 : BOOL;
  elapsed AT %QD1 : TIME;
END_VAR
  shot(IN := trigger, PT := T#30ms);
  q := shot.Q;
  elapsed := shot.ET;
END_PROGRAM

(* ---- cmp-057-tp-new-edge-starts-a-new-pulse.st ---- *)
PROGRAM Pulses
VAR
  trigger AT %IX0.0 : BOOL;
  shot : TP;
  q AT %QX0.0 : BOOL;
  elapsed AT %QD1 : TIME;
END_VAR
  shot(IN := trigger, PT := T#40ms);
  q := shot.Q;
  elapsed := shot.ET;
END_PROGRAM

(* ---- cmp-057-tp-not-retriggered.st ---- *)
PROGRAM Window
VAR
  t : TP;
  q AT %QX0.0 : BOOL;
END_VAR
  t(IN := TRUE, PT := T#50ms);
  q := t.Q;
END_PROGRAM

(* ---- cmp-057-tp-pulse-ignores-the-input-falling.st ---- *)
PROGRAM PulseTimer
VAR
  trigger AT %IX0.0 : BOOL;
  shot : TP;
  q AT %QX0.0 : BOOL;
END_VAR
  shot(IN := trigger, PT := T#50ms);
  q := shot.Q;
END_PROGRAM

(* ---- cmp-057-trunc-keeps-negative-and-large-values.st ---- *)
PROGRAM Truncate
VAR
  negative : REAL := -3.7;
  fraction : REAL := 0.9;
  large : REAL := 3.0E9;
  t0 AT %QD0 : REAL;
  t1 AT %QD1 : REAL;
  t2 AT %QD2 : REAL;
  t3 AT %QD3 : REAL;
END_VAR
  t0 := TRUNC(negative);
  t1 := TRUNC(fraction);
  t2 := TRUNC(large);
  t3 := TRUNC(0.0 - fraction);
END_PROGRAM

(* ---- cmp-057-trunc-truncates.st ---- *)
PROGRAM Convert
VAR
  r : REAL := 3.7;
  whole AT %QD0 : REAL;
END_VAR
  whole := TRUNC(r);
END_PROGRAM

(* ---- cmp-058-absf-and-negf-of-negative-and-zero-values.st ---- *)
PROGRAM Signs
VAR
  neg : REAL := -3.5;
  pos : REAL := 2.5;
  zero : REAL := 0.0;
  big : REAL := -1.0E30;
  q0 AT %QD0 : REAL;
  q1 AT %QD1 : REAL;
  q2 AT %QD2 : REAL;
  q3 AT %QD3 : REAL;
  q4 AT %QD4 : REAL;
  q5 AT %QD5 : REAL;
  q6 AT %QD6 : REAL;
  q7 AT %QD7 : REAL;
END_VAR
  q0 := ABSF(neg);
  q1 := ABSF(pos);
  q2 := ABSF(zero);
  q3 := ABSF(big);
  q4 := NEGF(pos);
  q5 := NEGF(neg);
  q6 := NEGF(zero);
  q7 := NEGF(big);
END_PROGRAM

(* ---- cmp-058-blink-alternates-on-and-off.st ---- *)
PROGRAM Lamp
VAR
  enable AT %IX0.0 : BOOL;
  flasher : BLINK;
  q AT %QX0.0 : BOOL;
END_VAR
  flasher(ENABLE := enable, T_ON := T#30ms, T_OFF := T#20ms);
  q := flasher.Q;
END_PROGRAM

(* ---- cmp-058-blink-starts-on-again-after-it-is-disabled.st ---- *)
PROGRAM Lamp
VAR
  enable AT %IX0.0 : BOOL;
  flasher : BLINK;
  q AT %QX0.0 : BOOL;
END_VAR
  flasher(ENABLE := enable, T_ON := T#30ms, T_OFF := T#20ms);
  q := flasher.Q;
END_PROGRAM

(* ---- cmp-058-copy-and-clear-string-functions.st ---- *)
PROGRAM Edit
VAR
  source : STRING[20] := 'hello';
  target : STRING[20] := 'xxxxxxxxxxxxxxxx';
  other : STRING[20] := 'abc';
  short : STRING[3] := 'zzz';
  l0 AT %QW0 : INT;
  l1 AT %QW1 : INT;
  l2 AT %QW2 : INT;
  l3 AT %QW3 : INT;
  same AT %QX8.0 : BOOL;
  kept AT %QX8.1 : BOOL;
END_VAR
  target := COPY(source, target);
  l0 := LEN(target);
  same := EQ_STRING(target, 'hello');
  other := CLEAR(other);
  l1 := LEN(other);
  short := COPY(source, short);
  l2 := LEN(short);
  kept := EQ_STRING(source, 'hello');
  l3 := LEN(source);
END_PROGRAM

(* ---- cmp-058-ctd-counts-below-zero.st ---- *)
PROGRAM CtdBelowZero
VAR
  cdIn AT %IX0.0 : BOOL;
  ldIn AT %IX0.1 : BOOL;
  c : CTD;
  q AT %QX0.0 : BOOL;
  cv AT %QW1 : INT;
END_VAR
  c(CD := cdIn, LD := ldIn, PV := 2);
  q := c.Q;
  cv := c.CV;
END_PROGRAM

(* ---- cmp-058-ctd-edge-during-load-is-not-counted.st ---- *)
PROGRAM CtdEdgeDuringLoad
VAR
  cdIn AT %IX0.0 : BOOL;
  ldIn AT %IX0.1 : BOOL;
  c : CTD;
  q AT %QX0.0 : BOOL;
  cv AT %QW1 : INT;
END_VAR
  c(CD := cdIn, LD := ldIn, PV := 3);
  q := c.Q;
  cv := c.CV;
END_PROGRAM

(* ---- cmp-058-ctd-edge-on-the-scan-load-is-released-counts.st ---- *)
PROGRAM CtdEdgeOnLoadRelease
VAR
  cdIn AT %IX0.0 : BOOL;
  ldIn AT %IX0.1 : BOOL;
  c : CTD;
  q AT %QX0.0 : BOOL;
  cv AT %QW1 : INT;
END_VAR
  c(CD := cdIn, LD := ldIn, PV := 3);
  q := c.Q;
  cv := c.CV;
END_PROGRAM

(* ---- cmp-058-ctd-stops-at-the-int-minimum.st ---- *)
PROGRAM CtdLowerLimit
VAR
  cdIn AT %IX0.0 : BOOL;
  ldIn AT %IX0.1 : BOOL;
  c : CTD;
  q AT %QX0.0 : BOOL;
  cv AT %QW1 : INT;
END_VAR
  c(CD := cdIn, LD := ldIn, PV := -32767);
  q := c.Q;
  cv := c.CV;
END_PROGRAM

(* ---- cmp-058-ctu-counts-to-preset.st ---- *)
PROGRAM Counter
VAR
  c : CTU;
  clk : BOOL;
  reached AT %QX0.0 : BOOL;
  value AT %QW1 : INT;
END_VAR
  clk := NOT clk;
  c(CU := clk, R := FALSE, PV := 3);
  reached := c.Q;
  value := c.CV;
END_PROGRAM

(* ---- cmp-058-ctu-edge-during-reset-is-not-counted.st ---- *)
PROGRAM CtuEdgeDuringReset
VAR
  cuIn AT %IX0.0 : BOOL;
  rIn AT %IX0.1 : BOOL;
  c : CTU;
  q AT %QX0.0 : BOOL;
  cv AT %QW1 : INT;
END_VAR
  c(CU := cuIn, R := rIn, PV := 1);
  q := c.Q;
  cv := c.CV;
END_PROGRAM

(* ---- cmp-058-ctu-edge-on-the-scan-reset-is-released-counts.st ---- *)
PROGRAM CtuEdgeOnResetRelease
VAR
  cuIn AT %IX0.0 : BOOL;
  rIn AT %IX0.1 : BOOL;
  c : CTU;
  q AT %QX0.0 : BOOL;
  cv AT %QW1 : INT;
END_VAR
  c(CU := cuIn, R := rIn, PV := 1);
  q := c.Q;
  cv := c.CV;
END_PROGRAM

(* ---- cmp-058-ctu-held-input-counts-once.st ---- *)
PROGRAM CtuHeldInput
VAR
  cuIn AT %IX0.0 : BOOL;
  rIn AT %IX0.1 : BOOL;
  c : CTU;
  q AT %QX0.0 : BOOL;
  cv AT %QW1 : INT;
END_VAR
  c(CU := cuIn, R := rIn, PV := 3);
  q := c.Q;
  cv := c.CV;
END_PROGRAM

(* ---- cmp-058-ctu-stops-at-32767.st ---- *)
PROGRAM CtuUpperLimit
VAR
  cuIn AT %IX0.0 : BOOL;
  rIn AT %IX0.1 : BOOL;
  c : CTU;
  q AT %QX0.0 : BOOL;
  cv AT %QW1 : INT;
  first : BOOL := TRUE;
END_VAR
  (* CV is written once to start next to the limit: reaching 32767 by counting takes 65534 scans *)
  IF first THEN
    c.CV := 32766;
    first := FALSE;
  END_IF;
  c(CU := cuIn, R := rIn, PV := 5);
  q := c.Q;
  cv := c.CV;
END_PROGRAM

(* ---- cmp-058-ctu-with-a-negative-preset.st ---- *)
PROGRAM CtuNegativePreset
VAR
  cuIn AT %IX0.0 : BOOL;
  rIn AT %IX0.1 : BOOL;
  c : CTU;
  q AT %QX0.0 : BOOL;
  cv AT %QW1 : INT;
END_VAR
  c(CU := cuIn, R := rIn, PV := -3);
  q := c.Q;
  cv := c.CV;
END_PROGRAM

(* ---- cmp-058-ctud-counts-down-through-zero-and-back.st ---- *)
PROGRAM CtudThroughZero
VAR
  cuIn AT %IX0.0 : BOOL;
  cdIn AT %IX0.1 : BOOL;
  c : CTUD;
  qu AT %QX0.0 : BOOL;
  qd AT %QX0.1 : BOOL;
  cv AT %QW1 : INT;
END_VAR
  c(CU := cuIn, CD := cdIn, R := FALSE, LD := FALSE, PV := -1);
  qu := c.QU;
  qd := c.QD;
  cv := c.CV;
END_PROGRAM

(* ---- cmp-058-ctud-load-beats-count-edges.st ---- *)
PROGRAM CtudLoadBeatsEdges
VAR
  cuIn AT %IX0.0 : BOOL;
  cdIn AT %IX0.1 : BOOL;
  rIn AT %IX0.2 : BOOL;
  ldIn AT %IX0.3 : BOOL;
  c : CTUD;
  qu AT %QX0.0 : BOOL;
  qd AT %QX0.1 : BOOL;
  cv AT %QW1 : INT;
END_VAR
  c(CU := cuIn, CD := cdIn, R := rIn, LD := ldIn, PV := 3);
  qu := c.QU;
  qd := c.QD;
  cv := c.CV;
END_PROGRAM

(* ---- cmp-058-ctud-reset-beats-count-edges.st ---- *)
PROGRAM CtudResetBeatsEdges
VAR
  cuIn AT %IX0.0 : BOOL;
  cdIn AT %IX0.1 : BOOL;
  rIn AT %IX0.2 : BOOL;
  ldIn AT %IX0.3 : BOOL;
  c : CTUD;
  qu AT %QX0.0 : BOOL;
  qd AT %QX0.1 : BOOL;
  cv AT %QW1 : INT;
END_VAR
  c(CU := cuIn, CD := cdIn, R := rIn, LD := ldIn, PV := 3);
  qu := c.QU;
  qd := c.QD;
  cv := c.CV;
END_PROGRAM

(* ---- cmp-058-ctud-reset-beats-load.st ---- *)
PROGRAM CtudResetBeatsLoad
VAR
  cuIn AT %IX0.0 : BOOL;
  cdIn AT %IX0.1 : BOOL;
  rIn AT %IX0.2 : BOOL;
  ldIn AT %IX0.3 : BOOL;
  c : CTUD;
  qu AT %QX0.0 : BOOL;
  qd AT %QX0.1 : BOOL;
  cv AT %QW1 : INT;
END_VAR
  c(CU := cuIn, CD := cdIn, R := rIn, LD := ldIn, PV := 3);
  qu := c.QU;
  qd := c.QD;
  cv := c.CV;
END_PROGRAM

(* ---- cmp-058-ctud-stops-at-32767.st ---- *)
PROGRAM CtudUpperLimit
VAR
  cuIn AT %IX0.0 : BOOL;
  cdIn AT %IX0.1 : BOOL;
  rIn AT %IX0.2 : BOOL;
  ldIn AT %IX0.3 : BOOL;
  c : CTUD;
  qu AT %QX0.0 : BOOL;
  qd AT %QX0.1 : BOOL;
  cv AT %QW1 : INT;
END_VAR
  c(CU := cuIn, CD := cdIn, R := rIn, LD := ldIn, PV := 32767);
  qu := c.QU;
  qd := c.QD;
  cv := c.CV;
END_PROGRAM

(* ---- cmp-058-ctud-up-and-down-edge-in-one-scan-cancel.st ---- *)
PROGRAM CtudBothEdges
VAR
  cuIn AT %IX0.0 : BOOL;
  cdIn AT %IX0.1 : BOOL;
  rIn AT %IX0.2 : BOOL;
  ldIn AT %IX0.3 : BOOL;
  c : CTUD;
  qu AT %QX0.0 : BOOL;
  qd AT %QX0.1 : BOOL;
  cv AT %QW1 : INT;
END_VAR
  c(CU := cuIn, CD := cdIn, R := rIn, LD := ldIn, PV := 5);
  qu := c.QU;
  qd := c.QD;
  cv := c.CV;
END_PROGRAM

(* ---- cmp-058-deadband-ignores-small-changes.st ---- *)
PROGRAM Quiet
VAR
  raw AT %ID0 : REAL;
  filter : DEADBAND;
  smooth AT %QD0 : REAL;
END_VAR
  filter(IN := raw, WIDTH := 1.0);
  smooth := filter.OUT;
END_PROGRAM

(* ---- cmp-058-deadband-with-negative-values.st ---- *)
PROGRAM Quiet
VAR
  raw AT %ID0 : REAL;
  filter : DEADBAND;
  smooth AT %QD0 : REAL;
END_VAR
  filter(IN := raw, WIDTH := 1.0);
  smooth := filter.OUT;
END_PROGRAM

(* ---- cmp-058-derivative-of-a-rising-and-falling-input.st ---- *)
PROGRAM Slope
VAR
  signal AT %ID0 : REAL;
  step : INT;
  d : DERIVATIVE;
  none : DERIVATIVE;
  rate AT %QD0 : REAL;
  guarded AT %QD1 : REAL;
END_VAR
  d(IN := signal, DT := 0.5);
  none(IN := signal, DT := 0.0);
  rate := d.OUT;
  guarded := none.OUT;
END_PROGRAM

(* ---- cmp-058-exp-ln-and-log-at-the-ends-of-their-ranges.st ---- *)
PROGRAM Exponentials
VAR
  q0 AT %QX0.0 : BOOL;
  q1 AT %QX0.1 : BOOL;
  q2 AT %QX0.2 : BOOL;
  q3 AT %QX0.3 : BOOL;
  q4 AT %QX0.4 : BOOL;
  q5 AT %QX0.5 : BOOL;
  q6 AT %QX0.6 : BOOL;
  q7 AT %QX0.7 : BOOL;
  q8 AT %QX1.0 : BOOL;
  q9 AT %QX1.1 : BOOL;
  q10 AT %QX1.2 : BOOL;
  q11 AT %QX1.3 : BOOL;
  q12 AT %QX1.4 : BOOL;
END_VAR
  q0 := ABS((EXP(-20.0) / 2.0611536E-9) - 1.0) < 1.0E-5;
  q1 := ABS((EXP(0.0)) - 1.0) < 1.0E-6;
  q2 := ABS((EXP(88.0) / 1.6516363E38) - 1.0) < 1.0E-5;
  q3 := EXP(100.0) > 3.0E38;
  q4 := EXP(-110.0) = 0.0;
  q5 := ABS((LN(1.0)) - 0.0) < 1.0E-6;
  q6 := ABS((LN(0.5)) - -0.6931471824645996) < 1.0E-6;
  q7 := ABS((LN(1.0E-40)) - -92.10340118408203) < 1.0E-4;
  q8 := LN(0.0) < -3.0E38;
  q9 := (LN(-1.0)) <> (LN(-1.0));
  q10 := ABS((LOG(100.0)) - 2.0) < 1.0E-6;
  q11 := ABS((LOG(0.001)) - -3.0) < 1.0E-6;
  q12 := ABS((LOG(1.0E30)) - 30.0) < 1.0E-5;
END_PROGRAM

(* ---- cmp-058-expt-integer-exponents-zero-and-negative.st ---- *)
PROGRAM Powers
VAR
  base : REAL := 5.0;
  minus_base : REAL := -3.0;
  zero : REAL := 0.0;
  three : REAL := 3.0;
  i : INT;
  sum : REAL;
  q0 AT %QD0 : REAL;
  q1 AT %QD1 : REAL;
  q2 AT %QD2 : REAL;
  q3 AT %QD3 : REAL;
  q4 AT %QD4 : REAL;
  q5 AT %QD5 : REAL;
  q6 AT %QD6 : REAL;
  q7 AT %QD7 : REAL;
  q8 AT %QD8 : REAL;
  q9 AT %QD9 : REAL;
END_VAR
  q0 := EXPT(2.0, 8.0);
  q1 := EXPT(base, zero);
  q2 := EXPT(minus_base, zero);
  q3 := EXPT(zero, zero);
  q4 := EXPT(2.0, -2.0);
  q5 := EXPT(minus_base, three);
  q6 := EXPT(minus_base, 2.0);
  q7 := EXPT(2, 10);
  q8 := EXPT(zero, three);
  FOR i := 1 TO 20 DO
    sum := sum + EXPT(2.0, three);
  END_FOR;
  q9 := sum;
END_PROGRAM

(* ---- cmp-058-expt-real-exponent-and-the-operator.st ---- *)
PROGRAM RealPowers
VAR
  q0 AT %QX0.0 : BOOL;
  q1 AT %QX0.1 : BOOL;
  q2 AT %QX0.2 : BOOL;
  q3 AT %QX0.3 : BOOL;
  q4 AT %QX0.4 : BOOL;
  q5 AT %QX0.5 : BOOL;
END_VAR
  q0 := ABS((EXPT(9.0, 0.5)) - 3.0) < 1.0E-5;
  q1 := ABS((EXPT(2.0, 0.5)) - 1.4142135381698608) < 1.0E-5;
  q2 := ABS((EXPT(10.0, -1.5)) - 0.03162277489900589) < 1.0E-6;
  q3 := EXPT(7.0, 2.5) = 7.0 ** 2.5;
  q4 := (EXPT(-8.0, 0.5)) <> (EXPT(-8.0, 0.5));
  q5 := ABS((EXPT(1.0, 1000.0)) - 1.0) < 1.0E-6;
END_PROGRAM

(* ---- cmp-058-f-trig-pulses-on-the-falling-edge.st ---- *)
PROGRAM Edges
VAR
  signal AT %IX0.0 : BOOL;
  fall : F_TRIG;
  seen AT %QX0.0 : BOOL;
END_VAR
  fall(CLK := signal);
  seen := fall.Q;
END_PROGRAM

(* ---- cmp-058-fifo-and-lifo-called-in-a-loop.st ---- *)
PROGRAM Loop
VAR
  i : INT;
  line : FIFO;
  pile : LIFO;
  line_count AT %QD0 : DINT;
  pile_count AT %QD1 : DINT;
  line_first AT %QD2 : DINT;
END_VAR
  FOR i := 1 TO 40 DO
    line(PUSH := (i MOD 2) = 1, DATA_IN := i, SIZE := 8);
    pile(PUSH := (i MOD 2) = 1, DATA_IN := i, SIZE := 8);
  END_FOR;
  line_count := line.COUNT;
  pile_count := pile.COUNT;
  line(POP := TRUE);
  line_first := line.DATA_OUT;
END_PROGRAM

(* ---- cmp-058-fifo-pop-of-an-empty-queue-does-nothing.st ---- *)
PROGRAM Empty
VAR
  line : FIFO;
  count AT %QD0 : DINT;
  empty AT %QX4.0 : BOOL;
END_VAR
  line(POP := TRUE);
  count := line.COUNT;
  empty := line.EMPTY;
END_PROGRAM

(* ---- cmp-058-fifo-returns-values-in-order.st ---- *)
PROGRAM Queue
VAR
  push AT %IX0.0 : BOOL;
  pop AT %IX0.1 : BOOL;
  item AT %ID1 : DINT;
  line : FIFO;
  first AT %QD0 : DINT;
  count AT %QD1 : DINT;
  empty AT %QX8.0 : BOOL;
END_VAR
  line(PUSH := push, POP := pop, DATA_IN := item, SIZE := 8);
  first := line.DATA_OUT;
  count := line.COUNT;
  empty := line.EMPTY;
END_PROGRAM

(* ---- cmp-058-fifo-size-above-its-capacity-is-limited-to-eight.st ---- *)
PROGRAM Overfill
VAR
  n : INT;
  line : FIFO;
  guard : DINT := 77;
  count AT %QD0 : DINT;
  full AT %QX4.0 : BOOL;
  neighbour AT %QD2 : DINT;
END_VAR
  n := n + 1;
  line(PUSH := (n MOD 2) = 1, DATA_IN := n, SIZE := 16);
  count := line.COUNT;
  full := line.FULL;
  neighbour := guard;
END_PROGRAM

(* ---- cmp-058-hysteresis-switches-at-its-thresholds.st ---- *)
PROGRAM Thermostat
VAR
  level AT %ID0 : REAL;
  band : HYSTERESIS;
  q AT %QX0.0 : BOOL;
END_VAR
  band(IN := level, HIGH := 8.0, LOW := 3.0);
  q := band.Q;
END_PROGRAM

(* ---- cmp-058-hysteresis-with-negative-thresholds.st ---- *)
PROGRAM Cold
VAR
  level AT %ID0 : REAL;
  band : HYSTERESIS;
  q AT %QX0.0 : BOOL;
END_VAR
  band(IN := level, HIGH := -2.0, LOW := -6.0);
  q := band.Q;
END_PROGRAM

(* ---- cmp-058-integral-accumulates-resets-and-follows-a-negative-input.st ---- *)
PROGRAM Accumulator
VAR
  rate AT %ID0 : REAL;
  clear AT %IX8.0 : BOOL;
  total : INTEGRAL;
  out AT %QD0 : REAL;
END_VAR
  total(IN := rate, DT := 0.5, RESET := clear);
  out := total.OUT;
END_PROGRAM

(* ---- cmp-058-inverse-trigonometric-functions-at-their-boundaries.st ---- *)
PROGRAM InverseAngles
VAR
  q0 AT %QX0.0 : BOOL;
  q1 AT %QX0.1 : BOOL;
  q2 AT %QX0.2 : BOOL;
  q3 AT %QX0.3 : BOOL;
  q4 AT %QX0.4 : BOOL;
  q5 AT %QX0.5 : BOOL;
  q6 AT %QX0.6 : BOOL;
  q7 AT %QX0.7 : BOOL;
  q8 AT %QX1.0 : BOOL;
  q9 AT %QX1.1 : BOOL;
  q10 AT %QX1.2 : BOOL;
  q11 AT %QX1.3 : BOOL;
  q12 AT %QX1.4 : BOOL;
  q13 AT %QX1.5 : BOOL;
  q14 AT %QX1.6 : BOOL;
  q15 AT %QX1.7 : BOOL;
END_VAR
  q0 := ABS((ASIN(1.0)) - 1.5707963705062866) < 1.0E-6;
  q1 := ABS((ASIN(-1.0)) - -1.5707963705062866) < 1.0E-6;
  q2 := ABS((ACOS(1.0)) - 0.0) < 1.0E-6;
  q3 := ABS((ACOS(-1.0)) - 3.1415927410125732) < 1.0E-6;
  q4 := ABS((ACOS(-0.5)) - 2.094395160675049) < 1.0E-6;
  q5 := (ASIN(1.5)) <> (ASIN(1.5));
  q6 := ABS((ATAN(-1.0E10)) - -1.5707963705062866) < 1.0E-6;
  q7 := ABS((ATAN(1.0E-10) * 1.0E10) - 1.0) < 1.0E-4;
  q8 := ABS((ATAN2(1.0, -1.0)) - 2.356194496154785) < 1.0E-6;
  q9 := ABS((ATAN2(-1.0, -1.0)) - -2.356194496154785) < 1.0E-6;
  q10 := ABS((ATAN2(-1.0, 1.0)) - -0.7853981852531433) < 1.0E-6;
  q11 := ABS((ATAN2(1.0, 0.0)) - 1.5707963705062866) < 1.0E-6;
  q12 := ABS((ATAN2(-1.0, 0.0)) - -1.5707963705062866) < 1.0E-6;
  q13 := ABS((ATAN2(0.0, -1.0)) - 3.1415927410125732) < 1.0E-6;
  q14 := ABS((ATAN2(0.0, 0.0)) - 0.0) < 1.0E-6;
  q15 := ABS((ATAN2(3.0, 4.0)) - 0.6435011029243469) < 1.0E-6;
END_PROGRAM

(* ---- cmp-058-inverse-trigonometric-functions.st ---- *)
PROGRAM InverseTrigonometry
VAR
  asin_half AT %QX0.0 : BOOL;
  asin_neg AT %QX0.1 : BOOL;
  acos_half AT %QX0.2 : BOOL;
  acos_one AT %QX0.3 : BOOL;
  atan_one AT %QX0.4 : BOOL;
  atan_neg AT %QX0.5 : BOOL;
END_VAR
  asin_half := ABS(ASIN(0.5) - 0.5235988) < 0.001;
  asin_neg := ABS(ASIN(-0.5) + 0.5235988) < 0.001;
  acos_half := ABS(ACOS(0.5) - 1.0471976) < 0.001;
  acos_one := ABS(ACOS(1.0)) < 0.001;
  atan_one := ABS(ATAN(1.0) - 0.7853982) < 0.001;
  atan_neg := ABS(ATAN(-1.0) + 0.7853982) < 0.001;
END_PROGRAM

(* ---- cmp-058-lag-filter-approaches-the-input.st ---- *)
PROGRAM Smoothing
VAR
  raw AT %ID0 : REAL;
  lag : LAG_FILTER;
  smooth AT %QD0 : REAL;
END_VAR
  lag(IN := raw, GAIN := 0.5);
  smooth := lag.OUT;
END_PROGRAM

(* ---- cmp-058-lag-filter-with-a-negative-input.st ---- *)
PROGRAM Smoothing
VAR
  raw AT %ID0 : REAL;
  lag : LAG_FILTER;
  smooth AT %QD0 : REAL;
END_VAR
  lag(IN := raw, GAIN := 0.5);
  smooth := lag.OUT;
END_PROGRAM

(* ---- cmp-058-logarithmic-and-exponential-functions.st ---- *)
PROGRAM Logarithms
VAR
  ln_ten AT %QX0.0 : BOOL;
  ln_one AT %QX0.1 : BOOL;
  log_thousand AT %QX0.2 : BOOL;
  exp_one AT %QX0.3 : BOOL;
  exp_zero AT %QX0.4 : BOOL;
  exp_neg AT %QX0.5 : BOOL;
  sqrt_sixteen AT %QX0.6 : BOOL;
  sqrt_two AT %QX0.7 : BOOL;
END_VAR
  ln_ten := ABS(LN(10.0) - 2.3025851) < 0.001;
  ln_one := ABS(LN(1.0)) < 0.001;
  log_thousand := ABS(LOG(1000.0) - 3.0) < 0.001;
  exp_one := ABS(EXP(1.0) - 2.7182818) < 0.001;
  exp_zero := ABS(EXP(0.0) - 1.0) < 0.001;
  exp_neg := ABS(EXP(-1.0) - 0.3678794) < 0.001;
  sqrt_sixteen := ABS(SQRT(16.0) - 4.0) < 0.001;
  sqrt_two := ABS(SQRT(2.0) - 1.4142136) < 0.001;
END_PROGRAM

(* ---- cmp-058-mod-of-negative-operands.st ---- *)
PROGRAM Remainders
VAR
  a : INT := -7;
  b : INT := 3;
  c : INT := 7;
  d : INT := -3;
  big : DINT := -2147483647;
  q0 AT %QW0 : INT;
  q1 AT %QW1 : INT;
  q2 AT %QW2 : INT;
  q3 AT %QW3 : INT;
  q4 AT %QD2 : DINT;
END_VAR
  q0 := a MOD b;
  q1 := c MOD d;
  q2 := a MOD d;
  q3 := c MOD b;
  q4 := big MOD 10;
END_PROGRAM

(* ---- cmp-058-nand-and-nor-result-is-a-bool.st ---- *)
PROGRAM GateBits
VAR
  t : BOOL := TRUE;
  f : BOOL := FALSE;
  nand_true AT %QB0 : BYTE;
  nand_false AT %QB1 : BYTE;
  nor_true AT %QB2 : BYTE;
  nor_false AT %QB3 : BYTE;
END_VAR
  nand_true := BOOL_TO_USINT(NAND(f, t));
  nand_false := BOOL_TO_USINT(NAND(t, t));
  nor_true := BOOL_TO_USINT(NOR(f, f));
  nor_false := BOOL_TO_USINT(NOR(t, f));
END_PROGRAM

(* ---- cmp-058-nand-and-nor-truth-tables.st ---- *)
PROGRAM Gates
VAR
  t : BOOL := TRUE;
  f : BOOL := FALSE;
  nand00 AT %QX0.0 : BOOL;
  nand01 AT %QX0.1 : BOOL;
  nand10 AT %QX0.2 : BOOL;
  nand11 AT %QX0.3 : BOOL;
  nor00 AT %QX0.4 : BOOL;
  nor01 AT %QX0.5 : BOOL;
  nor10 AT %QX0.6 : BOOL;
  nor11 AT %QX0.7 : BOOL;
END_VAR
  IF NAND(f, f) THEN nand00 := TRUE; ELSE nand00 := FALSE; END_IF;
  IF NAND(f, t) THEN nand01 := TRUE; ELSE nand01 := FALSE; END_IF;
  IF NAND(t, f) THEN nand10 := TRUE; ELSE nand10 := FALSE; END_IF;
  IF NAND(t, t) THEN nand11 := TRUE; ELSE nand11 := FALSE; END_IF;
  IF NOR(f, f) THEN nor00 := TRUE; ELSE nor00 := FALSE; END_IF;
  IF NOR(f, t) THEN nor01 := TRUE; ELSE nor01 := FALSE; END_IF;
  IF NOR(t, f) THEN nor10 := TRUE; ELSE nor10 := FALSE; END_IF;
  IF NOR(t, t) THEN nor11 := TRUE; ELSE nor11 := FALSE; END_IF;
END_PROGRAM

(* ---- cmp-058-norm-x-and-scale-x-with-negative-ranges.st ---- *)
PROGRAM Scaling
VAR
  zero_range : REAL := 5.0;
  q0 AT %QD0 : REAL;
  q1 AT %QD1 : REAL;
  q2 AT %QD2 : REAL;
  q3 AT %QD3 : REAL;
  q4 AT %QD4 : REAL;
  q5 AT %QD5 : REAL;
  q6 AT %QD6 : REAL;
  q7 AT %QD7 : REAL;
  q8 AT %QD8 : REAL;
END_VAR
  q0 := NORM_X(-10.0, 0.0, 10.0);
  q1 := NORM_X(0.0, 5.0, 20.0);
  q2 := NORM_X(zero_range, zero_range, zero_range);
  q3 := NORM_X(0.0, 30.0, 20.0);
  q4 := NORM_X(-20.0, -15.0, -10.0);
  q5 := SCALE_X(-10.0, 0.5, 10.0);
  q6 := SCALE_X(0.0, 0.25, 20.0);
  q7 := SCALE_X(-5.0, 1.0, -1.0);
  q8 := SCALE_X(100.0, 0.0, 200.0);
END_PROGRAM

(* ---- cmp-058-pid-compact-integral-and-derivative-terms.st ---- *)
PROGRAM Controller
VAR
  actual AT %ID0 : REAL;
  slow : PID_Compact;
  fast : PID_Compact;
  integral_out AT %QD0 : REAL;
  derivative_out AT %QD1 : REAL;
  no_sample AT %QD2 : REAL;
  none : PID_Compact;
END_VAR
  slow(SP := 10.0, PV := 0.0, KP := 0.0, KI := 1.0, KD := 0.0, DT := 0.5, OUT_MIN := -100.0, OUT_MAX := 100.0);
  fast(SP := 10.0, PV := actual, KP := 0.0, KI := 0.0, KD := 1.0, DT := 0.5, OUT_MIN := -100.0, OUT_MAX := 100.0);
  none(SP := 10.0, PV := 4.0, KP := 2.0, KI := 1.0, KD := 1.0, OUT_MIN := -100.0, OUT_MAX := 100.0);
  integral_out := slow.OUT;
  derivative_out := fast.OUT;
  no_sample := none.OUT;
END_PROGRAM

(* ---- cmp-058-pid-compact-proportional-term-and-output-limits.st ---- *)
PROGRAM Controller
VAR
  actual AT %ID0 : REAL;
  pid : PID_Compact;
  out AT %QD0 : REAL;
END_VAR
  pid(SP := 10.0, PV := actual, KP := 2.0, KI := 0.0, KD := 0.0, DT := 0.1, OUT_MIN := -100.0, OUT_MAX := 100.0);
  out := pid.OUT;
END_PROGRAM

(* ---- cmp-058-pulse-one-pulse-per-rising-edge.st ---- *)
PROGRAM Strobe
VAR
  trigger AT %IX0.0 : BOOL;
  shot : PULSE;
  q AT %QX0.0 : BOOL;
END_VAR
  shot(TRIG := trigger, PT := T#30ms);
  q := shot.Q;
END_PROGRAM

(* ---- cmp-058-pwm-duty-cycle-and-disable.st ---- *)
PROGRAM Modulator
VAR
  run AT %IX0.0 : BOOL;
  third : PWM;
  never : PWM;
  always : PWM;
  whole : PWM;
  q AT %QX0.0 : BOOL;
  q_never AT %QX0.1 : BOOL;
  q_always AT %QX0.2 : BOOL;
  q_whole AT %QX0.3 : BOOL;
END_VAR
  third(ENABLE := run, PERIOD := T#100ms, DUTY := 0.3);
  never(ENABLE := run, PERIOD := T#100ms, DUTY := 0.0);
  always(ENABLE := run, PERIOD := T#100ms, DUTY := 1.0);
  whole(ENABLE := run, PERIOD := T#100ms, DUTY := 1);
  q := third.Q;
  q_never := never.Q;
  q_always := always.Q;
  q_whole := whole.Q;
END_PROGRAM

(* ---- cmp-058-pwm-fractional-on-time.st ---- *)
PROGRAM Modulator
VAR
  run AT %IX0.0 : BOOL;
  slow : PWM;
  q AT %QX0.0 : BOOL;
END_VAR
  slow(ENABLE := run, PERIOD := T#1000ms, DUTY := 0.0305);
  q := slow.Q;
END_PROGRAM

(* ---- cmp-058-pwm-zero-period-is-always-off.st ---- *)
PROGRAM Modulator
VAR
  run AT %IX0.0 : BOOL;
  none : PWM;
  q AT %QX0.0 : BOOL;
END_VAR
  none(ENABLE := run, PERIOD := T#0ms, DUTY := 0.5);
  q := none.Q;
END_PROGRAM

(* ---- cmp-058-r-trig-one-pulse-per-edge.st ---- *)
PROGRAM Edges
VAR
  r : R_TRIG;
  x : BOOL;
  pulses AT %QW0 : INT;
END_VAR
  x := NOT x;
  r(CLK := x);
  IF r.Q THEN
    pulses := pulses + 1;
  END_IF;
END_PROGRAM

(* ---- cmp-058-ramp-real-limits-the-rate-up-and-down.st ---- *)
PROGRAM Ramp
VAR
  target AT %ID0 : REAL;
  limiter : RAMP_REAL;
  smooth AT %QD0 : REAL;
END_VAR
  limiter(IN := target, RATE := 2.0);
  smooth := limiter.OUT;
END_PROGRAM

(* ---- cmp-058-sel-and-mux-with-negative-and-real-inputs.st ---- *)
PROGRAM Selection
VAR
  yes : BOOL := TRUE;
  no : BOOL := FALSE;
  last : INT := 2;
  beyond : INT := 3;
  below : INT := -1;
  q0 AT %QW0 : INT;
  q1 AT %QW1 : INT;
  q2 AT %QD1 : REAL;
  q3 AT %QW4 : INT;
  q4 AT %QW5 : INT;
  q5 AT %QW6 : INT;
  q6 AT %QW7 : INT;
  q7 AT %QD4 : REAL;
END_VAR
  q0 := SEL(no, -5, 7);
  q1 := SEL(yes, -5, 7);
  q2 := SEL(yes, 1.5, -2.5);
  q3 := MUX(0, -10, 20, 30);
  q4 := MUX(last, -10, 20, 30);
  q5 := MUX(beyond, -10, 20, 30);
  q6 := MUX(below, -10, 20, 30);
  q7 := MUX(1, -1.5, 2.5);
END_PROGRAM

(* ---- cmp-058-selection-and-limit-functions.st ---- *)
PROGRAM Functions
VAR
  root AT %QD0 : REAL;
  magnitude AT %QW2 : INT;
  largest AT %QW3 : INT;
  limited AT %QW4 : INT;
  chosen AT %QW5 : INT;
  muxed AT %QW6 : INT;
  smallest AT %QW7 : INT;
  rest AT %QW8 : INT;
END_VAR
  root := SQRT(16.0);
  magnitude := ABS(5);
  largest := MAX(3, 9);
  limited := LIMIT(0, 50, 10);
  chosen := SEL(TRUE, 1, 2);
  muxed := MUX(1, 10, 20, 30);
  smallest := MIN(4, 2);
  rest := 17 MOD 5;
END_PROGRAM

(* ---- cmp-058-shift-and-rotate-at-the-ends-of-their-widths.st ---- *)
PROGRAM Bits
VAR
  one : DWORD := 16#00000001;
  top : DWORD := 16#80000000;
  byte_value : BYTE := 16#81;
  word_value : WORD := 16#0001;
  all_ones : BYTE := 16#FF;
  q0 AT %QD0 : DWORD;
  q1 AT %QD1 : DWORD;
  q2 AT %QB8 : BYTE;
  q3 AT %QW5 : WORD;
  q4 AT %QB12 : BYTE;
  q5 AT %QD4 : DWORD;
  q6 AT %QB20 : BYTE;
  q7 AT %QB21 : BYTE;
END_VAR
  q0 := SHL(one, 31);
  q1 := SHR(top, 31);
  q2 := ROL(byte_value, 1);
  q3 := ROR(word_value, 1);
  q4 := SHL(all_ones, 4);
  q5 := ROL(top, 32);
  q6 := ROL(byte_value, 8);
  q7 := ROR(byte_value, 0);
END_PROGRAM

(* ---- cmp-058-sine-of-infinity-and-not-a-number.st ---- *)
PROGRAM Infinite
VAR
  big : REAL := 1.0E38;
  inf : REAL;
  nan : REAL;
  q0 AT %QX0.0 : BOOL;
  q1 AT %QX0.1 : BOOL;
  q2 AT %QX0.2 : BOOL;
  q3 AT %QX0.3 : BOOL;
  q4 AT %QX0.4 : BOOL;
  q5 AT %QX0.5 : BOOL;
END_VAR
  inf := big * big;
  nan := inf - inf;
  q0 := SIN(inf) <> SIN(inf);
  q1 := COS(0.0 - inf) <> COS(0.0 - inf);
  q2 := TAN(inf) <> TAN(inf);
  q3 := SIN(nan) <> SIN(nan);
  q4 := COS(nan) <> COS(nan);
  q5 := SIN(1.0) = SIN(1.0);
END_PROGRAM

(* ---- cmp-058-sqrt-zero-negative-subnormal-and-large-arguments.st ---- *)
PROGRAM SquareRoots
VAR
  big : REAL := 1.0E38;
  nan : REAL;
  q0 AT %QX0.0 : BOOL;
  q1 AT %QX0.1 : BOOL;
  q2 AT %QX0.2 : BOOL;
  q3 AT %QX0.3 : BOOL;
  q4 AT %QX0.4 : BOOL;
  q5 AT %QX0.5 : BOOL;
  q6 AT %QX0.6 : BOOL;
  q7 AT %QX0.7 : BOOL;
END_VAR
  nan := big * big;
  nan := nan - nan;
  q0 := ABS((SQRT(0.0)) - 0.0) < 1.0E-6;
  q1 := ABS((SQRT(-4.0)) - 0.0) < 1.0E-6;
  q2 := ABS((SQRT(16)) - 4.0) < 1.0E-6;
  q3 := ABS((SQRT(2.0)) - 1.4142135381698608) < 1.0E-6;
  q4 := ABS((SQRT(1.0E-40) * 1.0E20) - 1.0) < 1.0E-4;
  q5 := ABS((SQRT(2.0E38) / 1.0E19) - 1.4142135381698608) < 1.0E-5;
  q6 := ABS((SQRT(0.25)) - 0.5) < 1.0E-6;
  q7 := SQRT(nan) <> SQRT(nan);
END_PROGRAM

(* ---- cmp-058-sr-and-rs-dominance.st ---- *)
PROGRAM Latches
VAR
  s : SR;
  r : RS;
  set_wins AT %QX0.0 : BOOL;
  reset_wins AT %QX0.1 : BOOL;
END_VAR
  s(S1 := TRUE, R := TRUE);
  r(S := TRUE, R1 := TRUE);
  set_wins := s.Q1;
  reset_wins := r.Q1;
END_PROGRAM

(* ---- cmp-058-string-comparison-functions.st ---- *)
PROGRAM Compare
VAR
  apple : STRING[20] := 'apple';
  banana : STRING[20] := 'banana';
  upper : STRING[20] := 'Apple';
  empty : STRING[20] := '';
  c0 AT %QB0 : SINT;
  c1 AT %QB1 : SINT;
  c2 AT %QB2 : SINT;
  c3 AT %QB3 : SINT;
  c4 AT %QB4 : SINT;
  e0 AT %QX8.0 : BOOL;
  e1 AT %QX8.1 : BOOL;
  e2 AT %QX8.2 : BOOL;
  n0 AT %QX8.3 : BOOL;
  n1 AT %QX8.4 : BOOL;
  n2 AT %QX8.5 : BOOL;
END_VAR
  c0 := STRCMP(apple, banana);
  c1 := STRCMP(banana, apple);
  c2 := STRCMP(apple, apple);
  c3 := STRCMP(upper, apple);
  c4 := STRCMP(empty, empty);
  e0 := EQ_STRING(apple, 'apple');
  e1 := EQ_STRING(apple, banana);
  e2 := EQ_STRING(empty, empty);
  n0 := NE_STRING(apple, banana);
  n1 := NE_STRING(apple, 'apple');
  n2 := NE_STRING(upper, apple);
END_PROGRAM

(* ---- cmp-058-tof-holds-output.st ---- *)
PROGRAM Timer
VAR
  t : TOF;
  n : INT;
  q AT %QX0.0 : BOOL;
END_VAR
  n := n + 1;
  t(IN := n <= 2, PT := T#50ms);
  q := t.Q;
END_PROGRAM

(* ---- cmp-058-ton-delays-output.st ---- *)
PROGRAM Timer
VAR
  t : TON;
  q AT %QX0.0 : BOOL;
END_VAR
  t(IN := TRUE, PT := T#50ms);
  q := t.Q;
END_PROGRAM

(* ---- cmp-058-trigonometric-functions-of-negative-and-large-angles.st ---- *)
PROGRAM Angles
VAR
  q0 AT %QX0.0 : BOOL;
  q1 AT %QX0.1 : BOOL;
  q2 AT %QX0.2 : BOOL;
  q3 AT %QX0.3 : BOOL;
  q4 AT %QX0.4 : BOOL;
  q5 AT %QX0.5 : BOOL;
  q6 AT %QX0.6 : BOOL;
  q7 AT %QX0.7 : BOOL;
  q8 AT %QX1.0 : BOOL;
  q9 AT %QX1.1 : BOOL;
  q10 AT %QX1.2 : BOOL;
  q11 AT %QX1.3 : BOOL;
  q12 AT %QX1.4 : BOOL;
  q13 AT %QX1.5 : BOOL;
  q14 AT %QX1.6 : BOOL;
  q15 AT %QX1.7 : BOOL;
  q16 AT %QX2.0 : BOOL;
  q17 AT %QX2.1 : BOOL;
  q18 AT %QX2.2 : BOOL;
END_VAR
  q0 := ABS((SIN(100.0)) - -0.5063656568527222) < 1.0E-5;
  q1 := ABS((COS(1000.0)) - 0.5623790621757507) < 1.0E-5;
  q2 := ABS((SIN(-10000.0)) - 0.3056143820285797) < 1.0E-5;
  q3 := ABS((TAN(-0.5)) - -0.5463024973869324) < 1.0E-5;
  q4 := ABS((SIN(-0.5)) - -0.4794255495071411) < 1.0E-6;
  q5 := ABS((COS(-3.0)) - -0.9899924993515015) < 1.0E-6;
  q6 := ABS((SIN(3.1415927)) - 0.0) < 1.0E-6;
  q7 := ABS((COS(3.1415927)) - -1.0) < 1.0E-6;
  q8 := ABS((COS(6.2831855)) - 1.0) < 1.0E-6;
  q9 := ABS((SIN(0)) - 0.0) < 1.0E-6;
  q10 := ABS((TAN(0.7853982)) - 1.0) < 1.0E-5;
  q11 := ABS((SIN(100000.0)) - 0.03574879840016365) < 1.0E-5;
  q12 := ABS((SIN(1.0E6)) - -0.349993497133255) < 1.0E-5;
  q13 := ABS((COS(-1.0E6)) - 0.9367521405220032) < 1.0E-5;
  q14 := ABS((COS(1.0E9)) - 0.837887167930603) < 1.0E-5;
  q15 := ABS((SIN(1.0E11)) - 0.9981087446212769) < 1.0E-5;
  q16 := ABS((TAN(1.0E7)) - -0.46353083848953247) < 1.0E-4;
  q17 := ABS(SIN(3.0E38)) <= 1.0;
  q18 := ABS(TAN(3.0E38)) < 3.0E38;
END_PROGRAM

(* ---- cmp-058-trigonometric-functions.st ---- *)
PROGRAM Trigonometry
VAR
  sin_pos AT %QX0.0 : BOOL;
  sin_neg AT %QX0.1 : BOOL;
  cos_pos AT %QX0.2 : BOOL;
  cos_neg AT %QX0.3 : BOOL;
  tan_pos AT %QX0.4 : BOOL;
  tan_neg AT %QX0.5 : BOOL;
  sin_zero AT %QX0.6 : BOOL;
  cos_zero AT %QX0.7 : BOOL;
END_VAR
  sin_pos := ABS(SIN(1.0) - 0.8414710) < 0.001;
  sin_neg := ABS(SIN(-1.0) + 0.8414710) < 0.001;
  cos_pos := ABS(COS(1.0) - 0.5403023) < 0.001;
  cos_neg := ABS(COS(-1.0) - 0.5403023) < 0.001;
  tan_pos := ABS(TAN(1.0) - 1.5574077) < 0.001;
  tan_neg := ABS(TAN(-1.0) + 1.5574077) < 0.001;
  sin_zero := ABS(SIN(0.0)) < 0.001;
  cos_zero := ABS(COS(0.0) - 1.0) < 0.001;
END_PROGRAM

(* ---- cmp-058-uptime-follows-the-clock.st ---- *)
PROGRAM Clock
VAR
  up AT %QD0 : DINT;
  cycle_known AT %QX4.0 : BOOL;
  survived AT %QX4.1 : BOOL;
END_VAR
  up := UPTIME();
  cycle_known := CYCLE_TIME() >= 0;
  WATCHDOG_RESET();
  survived := TRUE;
END_PROGRAM
